(* CODESYS project Portal_robot.project

Project tree, tasks and I/O mapping:
  Device : LicOS-PAC-MC522, Unionscience Technology Group Co.,Ltd, order no. 50080156/50080256, version 3.5.18.50
      unmapped channels: ErrCode
    application Application
      libraries: Standard, 3.5.18.0 (System); CmpBitmapPool, * (System); ModbusFB, 4.3.0.0 (3S - Smart Software Solutions GmbH)
      task MainTask (cyclic, interval t#4ms, priority 0) calls PLC_PRG
      task StatisticTask (freewheeling, priority 3) calls STATISTIC
      task SoftMotion_PlanningTask (cyclic, interval t#2ms, priority 1) calls nothing
      image pool HMI_Image
      axis group AXIS_GROUP_XYZ: TRAFO.Kin_Gantry3, axes X, Y, Z
      Symbols
      FB/
        function block FB_MAGAZINE [ST]: FindBlank, UpdateErrorView, FindFreeSlot, UpdateTypeStatus
        function block FB_TWO_PALLET_SIMULATION [ST]
        function block FB_MOTION_MANAGER [ST]: UpdateErrorView
        function block FB_ALARM_MANAGER [ST]: DeactivateEvent, GetAlarmEffect, AddEvent, UpdateSource
        function block FB_SIMULATION_DYNAMIC_LIMITS [ST]
        function block FB_AXIS [ST]: UpdateErrorView
        function block FB_ALARM_HORN [ST]
        function F_GEOMETRY_EVENT [ST]
        function block FB_GRIPPER_SIMULATION [ST]: UpdateErrorView
        function block FB_MACHINE [ST]: UpdateErrorView
        function block FB_AXIS_GROUP [ST]: UpdateErrorView
        function block FB_GEOMETRY_CONTROL_SIMULATION [ST]
        function block FB_POINT_MANAGER [ST]: UpdateErrorView
        function block FB_ROBOT_MODBUS [ST]
        function block FB_DI_FILTER [ST]
        function block FB_GEOMETRY_CONTROL [ST]
        _ARCHIVE_LEGACY_MULTI_TYPE_HELPERS/
          function block FB_MAGAZINE_RETURN_BLANK_LEGACY [ST]
          function block FB_MAGAZINE_MULTI_TYPE_MAP_LEGACY [ST]
        FB_FAULT_INJECTOR/
          function block FB_ROBOT_FAULT_INJECTOR [ST]
          function block FB_MAGAZINE_FAULT_INJECTOR [ST]
          function block FB_CELL_SAFETY_FAULT_INJECTOR [ST]
          function block FB_CELL_FAULT_INJECTOR [ST]
          function block FB_AXIS_GROUP_FAULT_INJECTOR [ST]
          function block FB_POINT_FAULT_INJECTOR [ST]
          function block FB_GRIPPER_FAULT_INJECTOR [ST]
          function block FB_MACHINE_FAULT_INJECTOR [ST]
          function block FB_AXIS_FAULT_INJECTOR [ST]
        function block FB_ROBOT [ST]: UpdateErrorView
        _ARCHIVE_LEGACY_CELL_MANAGER/
          function block FB_CELL_MANAGER_LEGACY [ST]: UpdateErrorView, SelectMachine
        function F_GEOMETRY_SELECT_STATION [ST]
        function block FB_TWO_PALLET [ST]: IsSignalConfigurationValid, UpdateErrorView
        FB_STATISTIC/
          function block FB_CALCULATE [ST]
          function block FB_STATISTIC [ST]
        function block FB_MACHINE_SIMULATION [ST]: UpdateErrorView
        FB_MULTI_TYPE/
          function block FB_MULTI_TYPE_CONFIG_MANAGER [ST]: ApplyDistribution, RaiseWarning
        function F_GEOMETRY_FIRST_CALL [ST]
        FB_CELL_MANAGER/
          function block FB_CELL_MANAGER [ST]: IsMachineEligible, RaisePayloadRouteWarning, RunGeometryRoute, IsMachineCompatible, SelectMachineBeforeTake, PlanGeometry, UpdateErrorView, SelectMachineForUnload, UpdateGeometryWait, SelectMachineForHeldBlank, CanReturnHeldBlank
        function block FB_CELL_SAFETY [ST]: RaiseWarning
        function F_GEOMETRY_TAKE_DETAIL [ST]
      program PLC_PRG [ST]: ReadHmiInputs, ResetIoEmergencyStop, ReadHmiCommands, RunRobotModbus, RunRobot, RunTwoPallet, RunCellControl, RunTestControl, RunSignalTower, AppendIoEvent, RunMagazine, RunTwoPalletAxis, ReadIoEmergencyStop, RunMotion, RunGeometryControl, RunMachines, ApplyIoOutputOverrides, RunAlarms, ReadPhysicalInputs, RecordIoDiagnostics, PublishGeometryControl, SetApplicationDefaults, RunSafety, ReadIoOverrides, PublishHmi, IsHmiCommandFresh, WritePhysicalOutputs
      ST/
        ST_GRIPPER/
          data type E_GRIPPER_STATE
          data type ST_GRIPPER_DIAG
          data type ST_GRIPPER_COMMAND
          data type ST_GRIPPER_STATUS
          data type ST_GRIPPER_FAULT_REQUEST
          data type ST_GRIPPER_ERRORS
          data type ST_GRIPPER_ERROR
        ST_MULTI_TYPE/
          data type ST_MULTI_TYPE_CONFIG_STATUS
          data type ST_MULTI_TYPE_COMMAND
          data type ST_MULTI_TYPE_CONFIG
          data type ST_MULTI_TYPE_HMI
        ST_ALARM/
          data type ST_ALARM_EVENT
          data type E_ALARM_EFFECT
          data type ST_ALARM_STATUS
          data type ST_ALARM_COMMAND
          data type E_ALARM_SEVERITY
          data type ST_WARNING_EVENT
          data type ST_ALARM_SOURCE_DATA
          data type E_ALARM_SOURCE
        ST_HMI/
          data type ST_PHYSICAL_IO_EVENT
          data type ST_AXIS_HMI_COMMAND
          data type ST_HMI
          data type ST_ROBOT_HMI_STATUS
          data type E_HMI_MANUAL_REJECT
          data type ST_AXIS_HMI_STATUS
        ST_POINT/
          data type ST_POINT
          data type E_POINT_NAME
        ST_ROBOT/
          data type ST_ROBOT_MODBUS_CONFIG
          data type ST_ROBOT_STATUS
          data type E_ROBOT_MODBUS_EXECUTION_STATE
          data type E_ROBOT_MODBUS_CLIENT_STATE
          data type ST_ROBOT_MODBUS_STATUS
          data type ST_ROBOT_FAULT_STATUS
          data type ST_ROBOT_ERRORS
          data type ST_ROBOT_FAULT_REQUEST
          data type ST_ROBOT_DIAG
          data type E_ROBOT_STATE
          data type ST_ROBOT_COMMAND
          data type ST_ROBOT_ERROR
          data type E_ROBOT_ACTION
          data type E_ROBOT_CONTROL_MODE
        ST_CELL/
          data type ST_CELL_DIAG
          data type ST_CELL_ERROR
          data type ST_CELL_SAFETY_DIAG
          data type ST_CELL_SAFETY_ERRORS
          data type ST_CELL_CYCLE_STATUS
          data type ST_ENCLOSURE_DOOR_STATUS
          data type ST_CELL_ERRORS
          data type ST_CELL_COMMAND
          data type ST_BUTTON_STATION_IO_STATUS
          data type E_CELL_MANAGER_STATE
          data type ST_CELL_FAULT_REQUEST
          data type ST_CONTROL_CABINET_IO_STATUS
          data type ST_CELL_STATUS
          data type ST_CELL_SAFETY_STATUS
          data type ST_MPG_IO_STATUS
          data type ST_CELL_SAFETY_FAULT_REQUEST
          data type E_CELL_STATE
        ST_TEST/
          data type ST_TEST_OBSERVABILITY
          data type ST_TEST_SCENARIO_BUFFER
          data type E_CELL_TEST_ENVIRONMENT
          data type E_TEST_SPEED_PROFILE
        ST_AXIS_GROUP/
          data type ST_AXIS_GROUP_ERROR
          data type ST_AXIS_GROUP_ERRORS
          data type ST_AXIS_GROUP_COMMANDS
          data type ST_AXIS_GROUP
          data type ST_AXIS_GROUP_TIMEOUTS
          data type ST_AXIS_GROUP_FAULT_REQUEST
          data type ST_AXIS_GROUP_MOTION_PARAMS
          data type E_AXIS_GROUP_POWER_MODE
          data type E_AXIS_GROUP_STATE
          data type ST_AXIS_GROUP_STATUS
          data type E_MOTION_RESET_STATE
          data type ST_AXIS_GROUP_DIAGNOSTICS
        ST_MOTION_MANAGER/
          data type ST_MOTION_MANAGER_DIAG
          data type ST_MOTION_MANAGER_ERROR
          data type ST_MOTION_MANAGER_COMMAND
          data type E_MOTION_MANAGER_STATE
          data type ST_MOTION_MANAGER
          data type ST_MOTION_MANAGER_ERRORS
          data type ST_MOTION_MANAGER_STATUS
        ST_POINT_MANAGER/
          data type ST_POINT_MANAGER_DIAG
          data type ST_POINT_FAULT_REQUEST
          data type ST_POINT_MANAGER_COMMAND
          data type E_POINT_MANAGER_STATE
          data type ST_POINT_MANAGER_ERRORS
          data type ST_POINT_MANAGER
          data type ST_POINT_MANAGER_ERROR
          data type ST_POINT_MANAGER_STATUS
        ST_MACHINE/
          data type ST_MACHINE_COMMAND
          data type E_PART_TYPE
          data type E_PART_STATE
          data type ST_MACHINE_SIM_ERROR
          data type ST_MACHINE_SIM_ERRORS
          data type ST_MACHINE_ERRORS
          data type ST_MACHINE_POINTS
          data type E_MACHINE_OPERATION
          data type ST_MACHINE_SIM_DIAG
          data type ST_MACHINE_ERROR
          data type ST_MACHINE_RECIPE
          data type ST_MACHINE_TIMEOUTS
          data type E_MACHINE_STATE
          data type ST_MACHINE_DIAG
          data type ST_MACHINE_IO_COMMAND
          data type ST_MACHINE_FAULT_REQUEST
          data type ST_MACHINE_IO_STATUS
          data type E_MACHINE_POINTS
          data type ST_MACHINE_PUBLIC
        ST_STATISTIC/
          data type ST_STATISTIC
          data type ST_STATISTIC_MACHINE
          data type ST_STATISTIC_ROBOT
        ST_GEOMETRY_CONTROL/
          data type ST_GEOMETRY_CALL
          data type ST_GEOMETRY_REQUEST
          data type ST_GEOMETRY_MEMORY
          data type ST_GEOMETRY_STATUS
          data type ST_GEOMETRY_CONFIG
          data type ST_GEOMETRY_SIGNALS
          data type ST_GEOMETRY_EVENT
        ST_MAGAZINE/
          data type ST_TWO_PALLET_ERROR
          data type ST_MAGAZINE_ERROR
          data type ST_MAGAZINE_TYPE_STATUS
          data type ST_MAGAZINE_STATUS
          data type ST_TWO_PALLET_INPUT
          data type ST_TWO_PALLET_ERRORS
          data type ST_MAGAZINE_DIAG
          data type ST_TWO_PALLET_COMMAND
          data type ST_MAGAZINE_FAULT_REQUEST
          data type ST_TWO_PALLET_DIAG
          data type ST_MAGAZINE_ERRORS
          data type ST_MAGAZINE_COMMAND
          data type E_MAGAZINE_STATE
          ST_DETAIL/
            data type E_DETAIL_TYPE
            data type ST_DETAIL
          data type E_TWO_PALLET_STATE
          data type ST_TWO_PALLET_CONFIG
          data type ST_MAGAZINE_HMI_COMMAND
          data type ST_TWO_PALLET_STATUS
          data type ST_TWO_PALLET_STORE
          data type E_MAGAZINE_OPERATION
          data type ST_MAGAZINE_INVENTORY
          data type ST_TWO_PALLET_REQUEST
          data type ST_TWO_PALLET_OUTPUT
        ST_AXIS/
          data type ST_AXIS_DIAGNOSTICS
          data type ST_AXIS_MOTION_PARAMS
          data type E_AXIS_STATE
          data type ST_AXIS_TIMEOUTS
          data type ST_AXIS_ERROR_CODES
          data type ST_AXIS_FAULT_REQUEST
          data type ST_AXIS
          data type ST_AXIS_STATUS
          data type ST_AXIS_ERROR
          data type ST_AXIS_COMMANDS
        ST_FAULT_INJECTOR/
          data type ST_FAULT_INJECTION_STATUS
      program STATISTIC [ST]
      GVL/
        global variables GVL_MAGAZINE
        global variables GVL_ROBOT
        global variables GVL_MAGAZINE_AXIS
        global variables GVL_MACHINE
        global variables GVL_POINT_MANAGER
        global variables GVL_HMI
        global variables GVL_AXIS_GROUP
        global variables GVL_ROBOT_MODBUS
        global variables GVL_CELL_CONTROL
        global variables GVL_CELL_MANAGER
        global variables GVL_POINT
        global variables GVL_ALARM
        global variables GVL_STATISTIC
        global variables GVL_ROBOT_MODBUS_RETAIN
        global variables GVL_CELL_SAFETY_IO
        global variables GVL_GEOMETRY_CONTROL
        global variables GVL_TEST_IO
        global variables GVL_CELL_SETTINGS
        global variables GVL_DETAIL
        global variables GVL_AXIS
        global variables GVL_MULTI_TYPE
        global variables GVL_MOTION_MANAGER
        global variables GVL_PHYSICAL_IO
        global variables GVL_TWO_PALLET
    SoftMotion General Axis Pool
      Z : SM_Drive_Virtual, 3S - Smart Software Solutions GmbH, order no. 1805, version 4.0.0.0
          settings: wDriveID = 0; fSWMaxVelocity = 3300; fSWMaxAcceleration = 12000; fSWMaxDeceleration = 12000; fSWMaxJerk = 100000; fSWLimitPositive = 10000.0; fSWLimitNegative = -1000.0; bSWLimitEnable = TRUE
      X : SM_Drive_Virtual, 3S - Smart Software Solutions GmbH, order no. 1805, version 4.0.0.0
          settings: fSWMaxVelocity = 3300; fSWMaxAcceleration = 12000; fSWMaxDeceleration = 12000; fSWMaxJerk = 100000; fSWLimitPositive = 13000.0; fSWLimitNegative = -1000.0; bSWLimitEnable = TRUE
      Y : SM_Drive_Virtual, 3S - Smart Software Solutions GmbH, order no. 1805, version 4.0.0.0
          settings: wDriveID = 2; fSWMaxVelocity = 3300; fSWMaxAcceleration = 12000; fSWMaxDeceleration = 12000; fSWMaxJerk = 100000; fSWLimitPositive = 10000.0; fSWLimitNegative = -1000.0; bSWLimitEnable = TRUE
      Magazine_1 : SM_Drive_Virtual, 3S - Smart Software Solutions GmbH, order no. 1805, version 4.0.0.0
          settings: wDriveID = 3; fSWMaxVelocity = 3300; fSWMaxAcceleration = 12000; fSWMaxDeceleration = 12000; fSWMaxJerk = 100000; fSWLimitPositive = 13000.0; fSWLimitNegative = -1000.0; bSWLimitEnable = TRUE
      Magazine_2 : SM_Drive_Virtual, 3S - Smart Software Solutions GmbH, order no. 1805, version 4.0.0.0
          settings: wDriveID = 4; fSWMaxVelocity = 3300; fSWMaxAcceleration = 12000; fSWMaxDeceleration = 12000; fSWMaxJerk = 100000; fSWLimitPositive = 13000.0; fSWLimitNegative = -1000.0; bSWLimitEnable = TRUE
    LicOS_MQTT : Mqtt Brok Sub Pub, Unionscience Technology Group Co.,Ltd, order no. 50010000, version 02.00.00.01
    LicOS_MTCP : ModbusTCP Device, Unionscience Technology Group Co.,Ltd, order no. 50011000, version 03.00.00.01
    LicOS_MUDP : ModbusUDP Device, Unionscience Technology Group Co.,Ltd, order no. 50011100, version 03.00.00.01
    LicOS_MRTU : ModbusRTU Device, Unionscience Technology Group Co.,Ltd, order no. 50012000, version 03.00.00.01
    LicOS_NETC : UDP/TCP NetComm, Unionscience Technology Group Co.,Ltd, order no. 50015000, version 01.00.00.01
    LicOS_INTM : Interrupt Cfg Module, Unionscience Technology Group Co.,Ltd, order no. 20110000, version 01.00.00.01
        unmapped channels: ErrCode
  libraries: VisuSymbols, 4.1.0.0 (System)
  text list GlobalTextList
*)

// Device/Application/ST/ST_CELL/ST_CELL_DIAG
TYPE ST_CELL_DIAG :
STRUCT
	eState : E_CELL_STATE; // Текущее состояние автомата ячейки
	stWarning : ST_WARNING_EVENT; // Последнее предупреждение менеджера ячейки
END_STRUCT
END_TYPE

// Device/Application/ST/ST_ROBOT/ST_ROBOT_MODBUS_CONFIG
TYPE ST_ROBOT_MODBUS_CONFIG :
STRUCT
	aIpAddress        : ARRAY [0..3] OF BYTE; // IPv4 контроллера робота
	uiPort            : UINT := UINT#502; // TCP-порт Modbus
	uiUnitId          : UINT := UINT#1; // Unit ID в Modbus TCP
	tResponseTimeout  : TIME := T#500MS; // Ожидание ответа FC03/FC16
	tPollInterval     : TIME := T#50MS; // Период чтения обратной связи
	tHeartbeatTimeout : TIME := T#2S; // Максимальная пауза heartbeat робота
	tCommandTimeout   : TIME := T#600S; // Предельная длительность одной команды
END_STRUCT
END_TYPE

// Device/Application/ST/ST_MOTION_MANAGER/ST_MOTION_MANAGER_DIAG
TYPE ST_MOTION_MANAGER_DIAG :
STRUCT
	eState : E_MOTION_MANAGER_STATE; // Текущее состояние автомата движения
	stWarning : ST_WARNING_EVENT; // Последнее предупреждение менеджера движения
END_STRUCT
END_TYPE

// Device/Application/ST/ST_CELL/ST_CELL_ERROR
TYPE ST_CELL_ERROR :
STRUCT
	BOTH_GRIPPERS_OCCUPIED : BOOL; // Совместимый бит: диагностическая ошибка согласованности захватов
	ROBOT_ERROR            : BOOL; // Ошибка робота во время автоматического цикла
	MAGAZINE_ERROR         : BOOL; // Ошибка магазина во время операции
	MACHINE_ERROR          : BOOL; // Ошибка станка во время обслуживания
	GLOBAL_STOP            : BOOL; // Получена глобальная ошибка ячейки
END_STRUCT
END_TYPE

// Device/Application/ST/ST_POINT_MANAGER/ST_POINT_MANAGER_DIAG
TYPE ST_POINT_MANAGER_DIAG :
STRUCT
	eState       : E_POINT_MANAGER_STATE; // Текущее состояние автомата
	lrX_MinLimit : LREAL; // Минимально допустимая координата X
	lrY_MinLimit : LREAL; // Минимально допустимая координата Y
	lrZ_MinLimit : LREAL; // Минимально допустимая координата Z
	lrX_MaxLimit : LREAL; // Максимально допустимая координата X
	lrY_MaxLimit : LREAL; // Максимально допустимая координата Y
	lrZ_MaxLimit : LREAL; // Максимально допустимая координата Z
	xXLimitValid : BOOL; // Software limits оси X включены и образуют корректный диапазон
	xYLimitValid : BOOL; // Software limits оси Y включены и образуют корректный диапазон
	xZLimitValid : BOOL; // Software limits оси Z включены и образуют корректный диапазон
	stWarning    : ST_WARNING_EVENT; // Последнее предупреждение менеджера точек
END_STRUCT
END_TYPE

// Device/Application/ST/ST_CELL/ST_CELL_SAFETY_DIAG
TYPE ST_CELL_SAFETY_DIAG :
STRUCT
	stWarning : ST_WARNING_EVENT; // Отклонённые попытки открытия и сброса реле
END_STRUCT
END_TYPE

// Device/Application/ST/ST_CELL/ST_CELL_SAFETY_ERRORS
TYPE ST_CELL_SAFETY_ERRORS :
STRUCT
	dwErrorActive : DWORD; // Текущие отдельные Safety-причины
	dwErrorLast   : DWORD; // Последняя ненулевая маска для диагностики
	dwAlarmActive : DWORD; // Собственные аварии источника для общего журнала
END_STRUCT
END_TYPE

// Device/Application/ST/ST_CELL/ST_CELL_CYCLE_STATUS
TYPE ST_CELL_CYCLE_STATUS :
STRUCT
	eState              : E_CELL_MANAGER_STATE; // Состояние универсального автомата ячейки
	uiSelectedMachine   : UINT; // Зафиксированный целевой станок
	uiSelectedType      : UINT; // Тип заготовки текущего маршрута
	uiBlankPayloadType  : UINT; // Тип заготовки в первом захвате
	uiDetailPayloadType : UINT; // Тип готовой детали во втором захвате
	iTakeSlot           : SINT; // Зарезервированный слот взятия
	iPutSlot            : SINT; // Зарезервированный слот укладки
	xReturningBlank     : BOOL; // Выполняется возврат заготовки
	axMachineStartPending: ARRAY [1..3] OF BOOL; // Запуск нового цикла ещё подтверждается станком
	auiBlankCount       : ARRAY [1..3] OF UINT; // Заготовки по типам
	auiDetailCount      : ARRAY [1..3] OF UINT; // Готовые детали по типам
	auiFreeCount        : ARRAY [1..3] OF UINT; // Свободные слоты по типам
END_STRUCT
END_TYPE

// Device/Application/ST/ST_TEST/ST_TEST_OBSERVABILITY
TYPE ST_TEST_OBSERVABILITY :
STRUCT
	udiAppliedScenarioSeq : UDINT;
	uiCellState : UINT;
	uiRobotState : UINT;
	uiRobotAction : UINT;
	uiRobotPoint : UINT;
	uiActiveMagazine : UINT;
	uiMagazineState : UINT;
	uiMagazineOperation : UINT;
	uiTakeSlot : UINT;
	uiPutSlot : UINT;
	auiMachineState : ARRAY [1..3] OF UINT;
	auiMachineOperation : ARRAY [1..3] OF UINT;
	uiSelectedMachine : UINT;
	uiSelectedType : UINT;
	uiErrorSource : UINT;
	dwErrorCode : DWORD;
END_STRUCT
END_TYPE

// Device/Application/ST/ST_MACHINE/ST_MACHINE_COMMAND
TYPE ST_MACHINE_COMMAND :
STRUCT
	stIo    : ST_MACHINE_IO_COMMAND; // Команды исполнительным механизмам станка
	stRobot : ST_ROBOT_COMMAND; // Команда роботу от алгоритма станка
END_STRUCT
END_TYPE

// Device/Application/ST/ST_MACHINE/E_PART_TYPE
{attribute 'qualified_only'}
{attribute 'strict'}
TYPE E_PART_TYPE :
(
	UNKNOWN,
	DETAIL,
	PART
);
END_TYPE

// Device/Application/ST/ST_MACHINE/E_PART_STATE
{attribute 'qualified_only'}
{attribute 'strict'}
TYPE E_PART_STATE :
(
	UNKNOWN := 0,
    EMPTY   := 1,
    LOADED  := 2
);
END_TYPE

// Device/Application/ST/ST_POINT_MANAGER/ST_POINT_FAULT_REQUEST
TYPE ST_POINT_FAULT_REQUEST :
STRUCT
	xEnabled        : BOOL; // Глобальное разрешение диагностической инъекции
	xXOutOfLimit    : BOOL; // Импульс проверки точки с недопустимой координатой X
	xYOutOfLimit    : BOOL; // Импульс проверки точки с недопустимой координатой Y
	xZOutOfLimit    : BOOL; // Импульс проверки точки с недопустимой координатой Z
	xInvalidVelocity: BOOL; // Импульс проверки точки с недопустимой скоростью
END_STRUCT
END_TYPE

// Device/Application/ST/ST_ROBOT/ST_ROBOT_STATUS
TYPE ST_ROBOT_STATUS :
STRUCT
	xBusy             : BOOL; // Робот выполняет команду
	xDone             : BOOL; // Команда завершена
	xError            : BOOL; // Робот находится в ошибке
	xExternalError    : BOOL; // Робот остановлен ошибкой зависимого блока
	xPowerAllowed     : BOOL; // Кнопка включения или отключения приводов доступна
	xStopAllowed      : BOOL; // Кнопка контролируемой остановки доступна
	xResetAllowed     : BOOL; // Кнопка сброса ошибок робота и приводов доступна
	eCurrentPoint     : E_POINT_NAME; // Последняя достигнутая точка
	uiMagazineContext : UINT; // 0 вне рабочей зоны; 1..2 — магазин, в рабочей зоне которого находится робот
	xBlankAvailable   : BOOL; // В первом захвате находится заготовка
	xDetailAvailable  : BOOL; // Во втором захвате находится готовая деталь
	uiBlankPayloadType  : UINT; // Фактический тип заготовки, 0 — неизвестно
	uiDetailPayloadType : UINT; // Фактический тип детали, 0 — неизвестно
	xGripper1Open     : BOOL; // Первый захват открыт
	xGripper1Closed   : BOOL; // Первый захват закрыт
	xGripper2Open     : BOOL; // Второй захват открыт
	xGripper2Closed   : BOOL; // Второй захват закрыт
	xRotatedToBlank   : BOOL; // Захват повёрнут к заготовке
	xRotatedToDetail  : BOOL; // Захват повёрнут к готовой детали
END_STRUCT
END_TYPE

// Device/Application/ST/ST_ROBOT/E_ROBOT_MODBUS_EXECUTION_STATE
{attribute 'qualified_only'}
{attribute 'strict'}
TYPE E_ROBOT_MODBUS_EXECUTION_STATE :
(
	IDLE := 0,
	ACCEPTED := 1,
	BUSY := 2,
	DONE := 3,
	ERROR := 4,
	STOPPED := 5
);
END_TYPE

// Device/Application/ST/ST_CELL/ST_ENCLOSURE_DOOR_STATUS
TYPE ST_ENCLOSURE_DOOR_STATUS :
STRUCT
	xLocked        : BOOL; // Обратная связь замка: TRUE — замок закрыт
	xUnlockAllowed : BOOL; // PLC разрешает открыть замок
	xUnlockOutput  : BOOL; // Фактическая команда открытия замка
END_STRUCT
END_TYPE

// Device/Application/ST/ST_ROBOT/E_ROBOT_MODBUS_CLIENT_STATE
{attribute 'qualified_only'}
{attribute 'strict'}
TYPE E_ROBOT_MODBUS_CLIENT_STATE :
(
	DISABLED,
	CONNECTING,
	INITIAL_READ,
	INITIAL_READ_RELEASE,
	CLEAR_COMMAND,
	CLEAR_COMMAND_RELEASE,
	READY,
	WRITE_COMMAND,
	WRITE_COMMAND_RELEASE,
	READ_STATUS,
	READ_STATUS_RELEASE,
	RECONNECT_WAIT
);
END_TYPE

// Device/Application/ST/ST_MAGAZINE/ST_TWO_PALLET_ERROR
TYPE ST_TWO_PALLET_ERROR :
STRUCT
	DRIVE_ERROR : BOOL;
	SENSOR_CONTRADICTION : BOOL;
	CYLINDER_TIMEOUT : BOOL;
	MOTION_TIMEOUT : BOOL;
	LOGIC_ERROR : BOOL;
	SEQUENCE_INTERRUPTED : BOOL;
END_STRUCT
END_TYPE

// Device/Application/ST/ST_MOTION_MANAGER/ST_MOTION_MANAGER_ERROR
TYPE ST_MOTION_MANAGER_ERROR :
STRUCT
	POINT_INVALID : BOOL; // Целевая точка не прошла проверку
	GROUP_ERROR   : BOOL; // Группа осей завершила движение с ошибкой
	GLOBAL_STOP   : BOOL; // Получена глобальная ошибка ячейки
	START_TIMEOUT : BOOL; // Истекло ожидание проверки точки или старта группы
END_STRUCT
END_TYPE

// Device/Application/ST/ST_AXIS/ST_AXIS_DIAGNOSTICS
TYPE ST_AXIS_DIAGNOSTICS :
STRUCT
    iStep            : E_AXIS_STATE; // Текущий шаг автомата оси
    iLastErrorStep   : INT; // Шаг, на котором возникла последняя ошибка
    sStepName        : STRING[80]; // Текстовое имя текущего шага
    sWaitReason      : STRING[120]; // Причина ожидания на текущем шаге
    sErrorText       : STRING[120]; // Текст активной ошибки
    sWarningText     : STRING[120]; // Текст активного предупреждения
    stWarning        : ST_WARNING_EVENT; // Последнее предупреждение оси для общего журнала
    tStepElapsed     : TIME; // Время нахождения на текущем шаге
    tStepPreset      : TIME; // Допустимое время текущего шага
    xStepTimeout     : BOOL; // Превышено допустимое время шага
    udiActualErrorID : UDINT; // Код активной ошибки
    udiLastErrorID   : UDINT; // Код последней ошибки
END_STRUCT
END_TYPE

// Device/Application/ST/ST_CELL/ST_CELL_ERRORS
TYPE ST_CELL_ERRORS :
STRUCT
	dwErrorActive : DWORD; // Битовая маска активных ошибок
	dwErrorLast   : DWORD; // Битовая маска последних ошибок
	dwAlarmActive : DWORD; // Собственные аварии менеджера ячейки для общего журнала
	stErrorActive : ST_CELL_ERROR; // Расшифровка активных ошибок
	stErrorLast   : ST_CELL_ERROR; // Расшифровка последних ошибок
END_STRUCT
END_TYPE

// Device/Application/ST/ST_AXIS/ST_AXIS_MOTION_PARAMS
TYPE ST_AXIS_MOTION_PARAMS :
STRUCT
    lrTargetPosition : LREAL; // Целевая абсолютная позиция
    lrDistance       : LREAL; // Дистанция относительного перемещения
    lrHomePosition   : LREAL; // Координата домашней позиции
    lrVelocity       : LREAL; // Скорость движения
    lrAcceleration   : LREAL; // Ускорение
    lrDeceleration   : LREAL; // Замедление
    lrJerk           : LREAL; // Рывок
END_STRUCT
END_TYPE

// Device/Application/ST/ST_ROBOT/ST_ROBOT_MODBUS_STATUS
TYPE ST_ROBOT_MODBUS_STATUS :
STRUCT
	xConfigValid       : BOOL; // Параметры соединения прошли проверку PLC
	xConnected         : BOOL; // TCP-соединение установлено
	xCommunicationAlive: BOOL; // Получена свежая обратная связь и меняется heartbeat
	xStatusFresh       : BOOL; // После подключения успешно прочитан блок 1101..1117
	xControllerOn      : BOOL;
	xAutomaticMode     : BOOL;
	xRemoteEnabled     : BOOL;
	xDrivesEnabled     : BOOL;
	xHomed             : BOOL;
	xEmergencyStop     : BOOL;
	xRobotAlarm        : BOOL;
	xPositionValid     : BOOL;
	xSimulatorActive   : BOOL; // Бит 1108.9: подключён Python-симулятор, а не реальный SC-500
	xReady             : BOOL; // Итоговая готовность, пересчитанная PLC
	xBusy              : BOOL;
	xDone              : BOOL;
	xError             : BOOL; // Ошибка исполнения, робота или транспорта
	xCommandTimeout    : BOOL; // Робот не завершил принятую команду за лимит
	xResetBusy         : BOOL; // Передача Reset и подтверждение его снятия ещё выполняются
	xResetDone         : BOOL; // Reset подтверждён обратной связью и очищенной FC16
	xResetFailed       : BOOL; // Попытка сорвана/истекла; повтор только новым запросом
	uiAckSeq           : UINT;
	uiExecutionState   : UINT;
	uiResultCode       : UINT;
	uiActiveCommand    : UINT;
	uiCurrentPoint     : UINT;
	uiGripperStatus    : UINT;
	uiRobotHeartbeat   : UINT;
	uiStatusWord       : UINT;
	uiAlarmCode        : UINT;
	uiOperationPhase   : UINT;
	uiProtocolVersion  : UINT;
	lrActualX          : LREAL;
	lrActualY          : LREAL;
	lrActualZ          : LREAL;
	udiClientError     : UDINT;
	udiReadError       : UDINT;
	udiWriteError      : UDINT;
END_STRUCT
END_TYPE

// Device/Application/ST/ST_AXIS/E_AXIS_STATE
{attribute 'qualified_only'}
{attribute 'strict'}
TYPE E_AXIS_STATE :
(
	DISABLED,
	POWERING,
	POWERING_DOWN,
	READY,
	JOGGING,
	JOG_DECELERATING,
	HOMING,
	MOVE_ABSOLUTE,
	MOVE_RELATIVE,
	STOPPING,
	STOP_RELEASE,
	ERROR_RESET_MANAGER,
	RESET_AXIS_ERROR,
	RESET_RELEASE,
	RESET_FINISH
);
END_TYPE

// Device/Application/ST/ST_AXIS/ST_AXIS_TIMEOUTS
TYPE ST_AXIS_TIMEOUTS :
STRUCT
	xDisableOnError : BOOL := TRUE; // Отключать привод при логической ошибке
    tPowerFeedbackLossTimeout : TIME := T#500MS; // Потеря силовой готовности при сохраняющемся запросе питания
    tPowerTimeout   : TIME := T#5S; // Время ожидания включения или отключения питания
    tResetTimeout   : TIME := T#5S; // Время ожидания сброса ошибки
    tStopTimeout    : TIME := T#5S; // Время ожидания остановки
    tHomeTimeout    : TIME := T#30S; // Время ожидания поиска домашней позиции
    tMoveTimeout    : TIME := T#15S; // Время ожидания завершения перемещения
END_STRUCT
END_TYPE

// Device/Application/ST/ST_ALARM/ST_ALARM_EVENT
TYPE ST_ALARM_EVENT :
STRUCT
	udiSequence : UDINT; // Уникальный порядковый номер события
	eSeverity   : E_ALARM_SEVERITY; // Уровень события
	eEffect     : E_ALARM_EFFECT; // Фактическое воздействие события в момент фиксации
	eSource     : E_ALARM_SOURCE; // Механизм-источник события
	uiCode      : UINT; // Номер бита ошибки или код предупреждения
	xActive     : BOOL; // Событие ещё активно и требует внимания
END_STRUCT
END_TYPE

// Device/Application/ST/ST_POINT_MANAGER/ST_POINT_MANAGER_COMMAND
TYPE ST_POINT_MANAGER_COMMAND :
STRUCT
	xExecute : BOOL; // Команда проверки заданной точки
END_STRUCT
END_TYPE

// Device/Application/ST/ST_MOTION_MANAGER/ST_MOTION_MANAGER_COMMAND
TYPE ST_MOTION_MANAGER_COMMAND :
STRUCT 
	eTargetPoint : E_POINT_NAME; // Имя целевой точки
	xGlobalError : BOOL; // Глобальная ошибка ячейки
	xExecute     : BOOL; // Команда запуска движения
	xStop        : BOOL; // Штатная операторская остановка без формирования аварии
	xReset       : BOOL; // Команда сброса ошибки
	xMode        : BOOL; // TRUE: Modbus, FALSE: SoftMotion
END_STRUCT
END_TYPE

// Device/Application/ST/ST_AXIS_GROUP/ST_AXIS_GROUP_ERROR
TYPE ST_AXIS_GROUP_ERROR :
STRUCT
	ENABLE_ERROR          : BOOL; // Ошибка MC_GroupEnable
	POWER_ERROR           : BOOL; // Зарезервировано; питание осей контролируют FB_AXIS
	DISABLE_ERROR         : BOOL; // Ошибка MC_GroupDisable
	RESET_ERROR           : BOOL; // Ошибка MC_GroupReset
	MOVE_DIRECT_ERROR     : BOOL; // Ошибка MC_MoveDirectAbsolute
	MOVE_LINEAR_ERROR     : BOOL; // Ошибка MC_MoveLinearAbsolute
	HALT_ERROR            : BOOL; // Ошибка MC_GroupHalt
	STOP_ERROR            : BOOL; // Ошибка MC_GroupStop
	READ_POSITION_ERROR   : BOOL; // Ошибка чтения позиции группы
	READ_STATUS_ERROR     : BOOL; // Ошибка чтения статуса группы
	READ_GROUP_ERROR      : BOOL; // Ошибка чтения кода ошибки группы
	GROUP_ERROR_STOP      : BOOL; // Группа SoftMotion находится в ErrorStop
	SIMULATED_ERROR       : BOOL; // Тестовая ошибка Motion-FB, сформированная эмулятором
	OVERRIDE_ERROR        : BOOL; // Ошибка MC_GroupSetOverride
	STEP_TIMEOUT          : BOOL; // Превышено время выполнения шага
	INVALID_STATE         : BOOL; // Неизвестное состояние автомата
	POWER_PERMIT_READY    : BOOL; // Нет разрешения питания в готовности
	POWER_PERMIT_LOST     : BOOL; // Потеря разрешения питания в движении
END_STRUCT
END_TYPE

// Device/Application/ST/ST_AXIS_GROUP/ST_AXIS_GROUP_ERRORS
TYPE ST_AXIS_GROUP_ERRORS :
STRUCT
	dwMotionErrorLatched  : DWORD; // Защёлкнутые ошибки SoftMotion
	dwLogicalErrorLatched : DWORD; // Защёлкнутые логические ошибки
	dwLogicalErrorNew     : DWORD; // Новые логические ошибки текущего цикла
	dwMotionErrorNew      : DWORD; // Новые ошибки SoftMotion текущего цикла
	dwMotionErrorActive   : DWORD; // Активные ошибки блоков SoftMotion
	dwMotionErrorPrevious : DWORD; // Ошибки SoftMotion предыдущего цикла
	dwMotionErrorLast     : DWORD; // Последняя ненулевая маска SoftMotion
	dwLogicalErrorLast    : DWORD; // Последняя ненулеевая логическая маска
	dwAlarmActive         : DWORD; // Собственные аварии группы для общего журнала
	stErrorActive         : ST_AXIS_GROUP_ERROR; // Расшифровка активных ошибок
	stErrorLast           : ST_AXIS_GROUP_ERROR; // Расшифровка последних ошибок
END_STRUCT
END_TYPE

// Device/Application/ST/ST_CELL/ST_CELL_COMMAND
TYPE ST_CELL_COMMAND :
STRUCT
	stRobot          : ST_ROBOT_COMMAND; // Команда роботу от менеджера ячейки
	uiBlankPayloadType  : UINT; // Тип заготовки в первом захвате
	uiDetailPayloadType : UINT; // Тип готовой детали во втором захвате
	stMagazine       : ST_MAGAZINE_COMMAND; // Команда магазину
	axMachineExecute : ARRAY [1..3] OF BOOL; // Запуск обслуживания выбранного станка
END_STRUCT
END_TYPE

// Device/Application/ST/ST_AXIS/ST_AXIS_ERROR_CODES
TYPE ST_AXIS_ERROR_CODES :
STRUCT
    dwAxisErrorActual     : DWORD; // Текущие ошибки блоков SoftMotion
    dwAxisErrorLatched    : DWORD; // Защёлкнутые ошибки SoftMotion
    dwAxisError           : DWORD; // Общая активная маска ошибок оси
    dwAxisErrorLast       : DWORD; // Последняя ненулевая маска ошибок оси
    dwDriveAxisErrorID    : DWORD; // Код ошибки привода
    dwLogicalErrorLatched : DWORD; // Защёлкнутые логические ошибки
    dwLogicalError        : DWORD; // Общая активная маска логических ошибок
    dwLogicalErrorLast    : DWORD; // Последняя ненулевая маска логических ошибок
    dwWarningLatched      : DWORD; // Защёлкнутые предупреждения
    dwWarning             : DWORD; // Активные предупреждения
    dwAllError            : DWORD; // Сводная маска ошибок
    dwAlarmActive         : DWORD; // Собственные аварии оси для общего журнала
    stErrorActive         : ST_AXIS_ERROR; // Расшифровка активных ошибок
    stErrorLast           : ST_AXIS_ERROR; // Расшифровка последних ошибок
END_STRUCT
END_TYPE

// Device/Application/ST/ST_MAGAZINE/ST_MAGAZINE_ERROR
TYPE ST_MAGAZINE_ERROR :
STRUCT
	WRONG_OPERATION : BOOL; // Операция не может быть выбрана
	NO_BLANK        : BOOL; // В магазине нет доступной заготовки
	NO_FREE_SLOT    : BOOL; // В магазине нет свободного слота
	INVALID_SLOT    : BOOL; // Номер слота находится вне матрицы
	SLOT_CONTENT    : BOOL; // Содержимое выбранного слота не соответствует операции
	ROBOT_ERROR     : BOOL; // Робот завершил команду с ошибкой
	GLOBAL_STOP     : BOOL; // Получена глобальная ошибка ячейки
	GEOMETRY_ERROR  : BOOL; // Геометрия магазина задана неверно
END_STRUCT
END_TYPE

// Device/Application/ST/ST_GRIPPER/E_GRIPPER_STATE
{attribute 'qualified_only'}
{attribute 'strict'}
TYPE E_GRIPPER_STATE :
(
	IDLE,
    EXECUTE,
    DONE,
    ERROR
);
END_TYPE

// Device/Application/ST/ST_ALARM/E_ALARM_EFFECT
TYPE E_ALARM_EFFECT :
(
	GLOBAL_STOP, // Аварийный останов всей ячейки
	ROBOT_STOP, // Останов робота и текущего взаимодействия с оборудованием
	EQUIPMENT_STOP, // Останов только владельца аварии
	WARNING // Информационное предупреждение без останова
);
END_TYPE

// Device/Application/ST/ST_ROBOT/ST_ROBOT_FAULT_STATUS
TYPE ST_ROBOT_FAULT_STATUS :
STRUCT
	stRobot   : ST_FAULT_INJECTION_STATUS; // Локальная ошибка автомата робота
	stGripper : ST_FAULT_INJECTION_STATUS; // Неисправности виртуального захвата
	stPoint   : ST_FAULT_INJECTION_STATUS; // Ошибки проверки точки движения
END_STRUCT
END_TYPE

// Device/Application/ST/ST_ALARM/ST_ALARM_STATUS
TYPE ST_ALARM_STATUS :
STRUCT
	uiActiveAlarmCount   : UINT; // Число активных аварий
	uiActiveWarningCount : UINT; // Число активных предупреждений
	uiActiveEventCount   : UINT; // Общее число активных событий
	uiHistoryCount       : UINT; // Число записей в журнале
	xAlarmActive         : BOOL; // Есть хотя бы одна активная авария
	xWarningActive       : BOOL; // Есть хотя бы одно активное предупреждение
END_STRUCT
END_TYPE

// Device/Application/ST/ST_MAGAZINE/ST_MAGAZINE_TYPE_STATUS
TYPE ST_MAGAZINE_TYPE_STATUS :
STRUCT
	aiBlankSlot    : ARRAY [1..3] OF SINT; // Первая заготовка каждого типа
	aiFreeSlot     : ARRAY [1..3] OF SINT; // Первый свободный слот каждого типа
	auiBlankCount  : ARRAY [1..3] OF UINT; // Количество заготовок каждого типа
	auiDetailCount : ARRAY [1..3] OF UINT; // Количество готовых деталей каждого типа
	auiFreeCount   : ARRAY [1..3] OF UINT; // Количество свободных слотов каждого типа
END_STRUCT
END_TYPE

// Device/Application/ST/ST_CELL/ST_BUTTON_STATION_IO_STATUS
TYPE ST_BUTTON_STATION_IO_STATUS :
STRUCT
	xEmergencyStopPressed : BOOL; // Нормализованный вход: TRUE — грибок нажат
	xButtonPressed        : BOOL; // Нормализованный вход кнопки открытия замка
	xButtonLightOn        : BOOL; // Фактический выход подсветки кнопки
END_STRUCT
END_TYPE

// Device/Application/ST/ST_MACHINE/ST_MACHINE_SIM_ERROR
TYPE ST_MACHINE_SIM_ERROR :
STRUCT
	MACHINE_ALARM : BOOL; // Активна имитация аварии станка
	DOOR_FAULT    : BOOL; // Ошибка механизма двери
	CHUCK_FAULT   : BOOL; // Ошибка механизма патрона
END_STRUCT
END_TYPE

// Device/Application/ST/ST_GRIPPER/ST_GRIPPER_DIAG
TYPE ST_GRIPPER_DIAG :
STRUCT
	eState        : E_GRIPPER_STATE; // Текущее состояние автомата
	eActiveAction : E_ROBOT_ACTION; // Выполняемое действие захвата
	stWarning     : ST_WARNING_EVENT; // Последнее предупреждение захвата
END_STRUCT
END_TYPE

// Device/Application/ST/ST_HMI/ST_PHYSICAL_IO_EVENT
TYPE ST_PHYSICAL_IO_EVENT :
STRUCT
    udiSequence : UDINT;
    uliTimeMs : ULINT; // Монотонное время от старта приложения, без переполнения TIME
    usiDirection : USINT; // 1 DI; 2 DO
    uiIndex : UINT; // DI 1..84; DO 1..50, index из карты I/O
    usiKind : USINT; // 1 клемма DI; 2 вход программы; 3 DO; 4 подмена DI; 5/6 снять DI; 7 ручной DO; 8/9 возврат DO оператором/программе
    xOld : BOOL;
    xNew : BOOL;
END_STRUCT
END_TYPE

// Device/Application/ST/ST_MAGAZINE/ST_MAGAZINE_STATUS
TYPE ST_MAGAZINE_STATUS :
STRUCT
	xEnabled         : BOOL; // Магазин включен в работу
	xDisablePending  : BOOL; // Отключение выполнится после выхода робота и завершения операции
	xPowerAllowed    : BOOL; // Команда включения/отключения может быть принята
	xEnableSequenceAllowed : BOOL; // PLC разрешает ввести подготовленный магазин в автомат
	xEnableCheckRobotReady : BOOL; // Диагностика готовности роботной операции; не блокирует включение
	xEnableCheckRobotReleased : BOOL; // Диагностика положения робота; не блокирует включение
	xEnableCheckNoError : BOOL; // Нет ошибок магазина и глобальных ошибок ячейки
	xEnableCheckContent : BOOL; // Содержимое кассеты допускает полезную операцию
	xEnableCheckGeometry : BOOL; // Матрица содержит от 1 до 120 активных слотов
	xFillAllowed     : BOOL; // Кнопка заполнения магазина заготовками доступна
	xClearAllowed    : BOOL; // Кнопка очистки магазина доступна
	xEditAllowed     : BOOL; // Содержимое разрешено менять только у выключенного магазина
	xPitchEditAllowed : BOOL; // Общий шаг X/Y можно менять только при выключенных обоих магазинах
	xReady 			 : BOOL; // Магазин готов принять команду
	xBusy  			 : BOOL; // Выполняется операция магазина
	xDone  			 : BOOL; // Операция магазина завершена
	xError          : BOOL; // Магазин находится в ошибке
	xRobotStopRequired : BOOL; // Ошибка магазина требует зависимой аварии робота
	xOutBlank        : BOOL; // В магазине не осталось свободных заготовок
	xOutFreeSlot     : BOOL; // В магазине не осталось свободных слотов
	xCanTake         : BOOL; // Операция TAKE доступна по содержимому магазина
	xCanPut          : BOOL; // Операция PUT доступна по содержимому магазина
	xCanChange       : BOOL; // Операция CHANGE доступна по содержимому магазина
	xCanEnable       : BOOL; // Содержимое позволяет взять/положить груз; не блокирует включение
	xFinished        : BOOL; // Палета завершена; защёлка до смены/правки её рабочего содержимого
	udiProducedPartsTotal : UDINT; // Подтверждённые укладки готовой детали с момента запуска PLC
	uiMagazineId    : UINT; // 1 или 2
	iCurrentBlank    : SINT; // Минимальный номер заготовки в матрице
	iCurrentFreeSlot : SINT; // Минимальный номер свободного слота в матрице
	iSelectedBlank   : SINT; // Номер заготовки, выбранной для текущей операции
	iSelectedFreeSlot: SINT; // Номер свободного слота, выбранного для текущей операции
	eGrantedOperation: E_MAGAZINE_OPERATION; // Доступная операция по текущему состоянию магазина
	eActualOperation : E_MAGAZINE_OPERATION; // Выполняемая операция магазина
	stTypeStatus     : ST_MAGAZINE_TYPE_STATUS; // Содержимое кассеты по типам
END_STRUCT
END_TYPE

// Device/Application/ST/ST_MULTI_TYPE/ST_MULTI_TYPE_CONFIG_STATUS
TYPE ST_MULTI_TYPE_CONFIG_STATUS :
STRUCT
	xMagazineConfigAllowed   : BOOL; // Типы и распределение слотов можно менять
	xTypeCountAllowed        : BOOL; // Количество типов можно менять с применением шаблона
	axMachineTypeAllowed     : ARRAY [1..3] OF BOOL; // Назначение типа конкретному станку разрешено
	xConfigurationValid      : BOOL; // Конфигурация пригодна для автоматического цикла
	uiActiveSlotCount        : UINT; // Число слотов активной матрицы
	stWarning                : ST_WARNING_EVENT; // Последняя отклонённая команда конфигурации
END_STRUCT
END_TYPE

// Device/Application/ST/ST_MACHINE/ST_MACHINE_SIM_ERRORS
TYPE ST_MACHINE_SIM_ERRORS :
STRUCT
	dwErrorActive : DWORD; // Битовая маска активных ошибок
	dwErrorLast   : DWORD; // Битовая маска последних ошибок
	stErrorActive : ST_MACHINE_SIM_ERROR; // Расшифровка активных ошибок
	stErrorLast   : ST_MACHINE_SIM_ERROR; // Расшифровка последних ошибок
END_STRUCT
END_TYPE

// Device/Application/ST/ST_MAGAZINE/ST_TWO_PALLET_INPUT
TYPE ST_TWO_PALLET_INPUT :
STRUCT
	xIoMapped : BOOL; // Подтверждается наладчиком после привязки и проверки физических I/O
	xLiftDown : BOOL;
	xLiftUp : BOOL;
	xLockIn : BOOL;
	xLockOut : BOOL;
	xStopIn : BOOL;
	xStopOut : BOOL;
	xLimitNegative : BOOL;
	xLimitPositive : BOOL;
	xHomeSensor : BOOL; // Только датчик каретки, не палет
	xAxisBound : BOOL;
	xPowered : BOOL;
	xHomed : BOOL;
	xStandstill : BOOL;
	xDriveError : BOOL;
	xMotionDone : BOOL;
	lrPosition : LREAL;
END_STRUCT
END_TYPE

// Device/Application/ST/ST_ROBOT/ST_ROBOT_ERRORS
TYPE ST_ROBOT_ERRORS :
STRUCT
	dwErrorActive : DWORD; // Битовая маска активных ошибок
	dwErrorLast   : DWORD; // Битовая маска последних ошибок
	dwAlarmActive : DWORD; // Собственные аварии робота для общего журнала
	stErrorActive : ST_ROBOT_ERROR; // Расшифровка активных ошибок
	stErrorLast   : ST_ROBOT_ERROR; // Расшифровка последних ошибок
END_STRUCT
END_TYPE

// Device/Application/ST/ST_HMI/ST_AXIS_HMI_COMMAND
TYPE ST_AXIS_HMI_COMMAND :
STRUCT
	xJogPositive      : BOOL; // Удерживаемый Jog в положительном направлении
	xJogNegative      : BOOL; // Удерживаемый Jog в отрицательном направлении
	{attribute 'symbol' := 'read'}
	xHome             : BOOL; // Импульс поиска домашней позиции выбранной оси
	{attribute 'symbol' := 'read'}
	xMoveAbsolute     : BOOL; // Импульс абсолютного перемещения к lrTargetPosition
	{attribute 'symbol' := 'read'}
	xMoveRelative     : BOOL; // Импульс относительного перемещения на lrRelativeDistance
	lrTargetPosition  : LREAL; // Целевая абсолютная координата оси
	lrRelativeDistance : LREAL; // Подготовленная дистанция относительного движения
END_STRUCT
END_TYPE

// Device/Application/ST/ST_HMI/ST_HMI
TYPE ST_HMI :
STRUCT
	ActualX : LREAL; // Текущая координата X для существующей визуализации
	ActualY : LREAL; // Текущая координата Y для существующей визуализации
	ActualZ : LREAL; // Текущая координата Z для существующей визуализации
END_STRUCT
END_TYPE

// Device/Application/ST/ST_GEOMETRY_CONTROL/ST_GEOMETRY_CALL
TYPE ST_GEOMETRY_CALL :
STRUCT
	udiId : UDINT; // Не меняется от вызова до результата контроля
	uiMachine : UINT;
	uiProductType : UINT;
	uiStation : UINT; // 0 до автоматического выбора свободного ГК
	xForced : BOOL;
	uiState : UINT; // 1 вызван, 2 в захвате/ожидание, 3 доставка, 4 на ГК, 5 в магазине, 6 отменён, 7 прерван, 8 изъят
	uiReason : UINT; // 1 заняты оба ГК, 2 нет доступного ГК, 3 отключён, 4 авария, 5 перезапуск/неопределённость
	uiMagazine : UINT;
	uiPallet : UINT;
	uiSlot : UINT;
END_STRUCT
END_TYPE

// Device/Application/ST/ST_STATISTIC/ST_STATISTIC
TYPE ST_STATISTIC :
STRUCT
	stMachineStat 		: ST_STATISTIC_MACHINE;
	stRobotStat 		: ST_STATISTIC_ROBOT;
END_STRUCT
END_TYPE

// Device/Application/ST/ST_ROBOT/ST_ROBOT_FAULT_REQUEST
TYPE ST_ROBOT_FAULT_REQUEST :
STRUCT
	xEnabled     : BOOL; // Глобальное разрешение диагностической инъекции
	xWrongAction : BOOL; // Импульс недопустимого действия робота
	stGripper : ST_GRIPPER_FAULT_REQUEST; // Неисправности виртуального захвата
	stPoint   : ST_POINT_FAULT_REQUEST; // Ошибки проверки точки движения
END_STRUCT
END_TYPE

// Device/Application/ST/ST_MACHINE/ST_MACHINE_ERRORS
TYPE ST_MACHINE_ERRORS :
STRUCT
	dwErrorActive : DWORD; // Битовая маска активных ошибок
	dwErrorLast   : DWORD; // Битовая маска последних ошибок
	dwAlarmActive : DWORD; // Собственные аварии станка для общего журнала
	stErrorActive : ST_MACHINE_ERROR; // Расшифровка активных ошибок
	stErrorLast   : ST_MACHINE_ERROR; // Расшифровка последних ошибок
END_STRUCT
END_TYPE

// Device/Application/ST/ST_MAGAZINE/ST_TWO_PALLET_ERRORS
TYPE ST_TWO_PALLET_ERRORS :
STRUCT
	dwErrorActive : DWORD;
	dwErrorLast : DWORD;
	dwAlarmActive : DWORD;
	stErrorActive : ST_TWO_PALLET_ERROR;
	stErrorLast : ST_TWO_PALLET_ERROR;
END_STRUCT
END_TYPE

// Device/Application/ST/ST_ROBOT/ST_ROBOT_DIAG
TYPE ST_ROBOT_DIAG :
STRUCT
	eState        : E_ROBOT_STATE; // Текущее состояние автомата робота
	eActiveAction : E_ROBOT_ACTION; // Выполняемое действие робота
	eActivePoint  : E_POINT_NAME; // Целевая точка текущего движения
	stWarning     : ST_WARNING_EVENT; // Последнее предупреждение робота
END_STRUCT
END_TYPE

// Device/Application/ST/ST_ALARM/ST_ALARM_COMMAND
TYPE ST_ALARM_COMMAND :
STRUCT
	xResetWarnings : BOOL; // Импульс сброса накопленных предупреждений
END_STRUCT
END_TYPE

// Device/Application/ST/ST_MOTION_MANAGER/E_MOTION_MANAGER_STATE
{attribute 'qualified_only'}
{attribute 'strict'}
TYPE E_MOTION_MANAGER_STATE :
(
	IDLE,
	VALIDATE,
	MOTION_SIM,
	MOTION_MODBUS,
	DONE,
	ERROR
);
END_TYPE

// Device/Application/ST/ST_MOTION_MANAGER/ST_MOTION_MANAGER
TYPE ST_MOTION_MANAGER :
STRUCT
	Command : ST_MOTION_MANAGER_COMMAND; // Команды менеджеру движения
	Status  : ST_MOTION_MANAGER_STATUS; // Рабочие статусы менеджера движения
	Diag    : ST_MOTION_MANAGER_DIAG; // Состояние автомата менеджера движения
	Error   : ST_MOTION_MANAGER_ERRORS; // Активные и последние ошибки
END_STRUCT
END_TYPE

// Device/Application/ST/ST_CELL/E_CELL_MANAGER_STATE
{attribute 'qualified_only'}
{attribute 'strict'}
TYPE E_CELL_MANAGER_STATE :
(
	IDLE,
	PLAN_TARGET,
	MAGAZINE_EXECUTE,
	RELEASE_MAGAZINE,
	ROUTE_TO_TARGET,
	RELEASE_ROBOT_COMMAND,
	WAIT_TARGET,
	SERVICE_TARGET,
	SELECT_FALLBACK,
	WAIT_MAGAZINE,
	ERROR,
	MACHINE_FAULT_STOP,
	PRESTART_IDENTIFY,
	WAIT_GRIPPER1_CONTENT,
	WAIT_GRIPPER1_TYPE,
	WAIT_GRIPPER2_CONTENT,
	WAIT_GRIPPER2_TYPE,
	WAIT_START_MACHINE,
	TEST_ABORT_STOP,
	GEOMETRY_WAIT_FREE,
	GEOMETRY_DELIVER,
	GEOMETRY_RELEASE_COMMAND
);
END_TYPE

// Device/Application/ST/ST_HMI/ST_ROBOT_HMI_STATUS
TYPE ST_ROBOT_HMI_STATUS :
STRUCT
	xDrivesPowered       : BOOL; // Все три привода фактически включены
	xDrivesOff           : BOOL; // Все три привода и группа фактически отключены
	xPowerTransitionActive : BOOL; // Выполняется последовательность включения или отключения
	xDrivesEnableAllowed : BOOL; // PLC разрешает включение приводов
	xDrivesDisableAllowed : BOOL; // PLC разрешает отключение приводов
	xResetAllowed        : BOOL; // PLC разрешает команду сброса ручного управления
	xStopAllowed         : BOOL; // PLC разрешает контролируемую остановку
	xPointsAllowed        : BOOL; // PLC разрешает переход к именованной точке
	xGripperAllowed       : BOOL; // PLC разрешает действие захвата
	xGripper1OpenAllowed  : BOOL;
	xGripper1CloseAllowed : BOOL;
	xGripper2OpenAllowed  : BOOL;
	xGripper2CloseAllowed : BOOL;
	xRotateToBlankAllowed : BOOL;
	xRotateToDetailAllowed : BOOL;
	xCommandBusy          : BOOL;
	uiActiveAction        : UINT;
	uiActivePoint         : UINT;
	eRejectReason         : E_HMI_MANUAL_REJECT; // Числовая причина недоступности команды
END_STRUCT
END_TYPE

// Device/Application/ST/ST_GRIPPER/ST_GRIPPER_COMMAND
TYPE ST_GRIPPER_COMMAND :
STRUCT
	xExecute : BOOL; // Команда запуска действия
	xReset   : BOOL; // Команда сброса ошибки
	eAction  : E_ROBOT_ACTION; // Требуемое действие захвата
	// Дискретный контракт исполнительных механизмов. Каждый BOOL задаёт
	// состояние своего механизма: 0 — закрыть/к заготовке, 1 — открыть/к детали.
	xGripper1Open   : BOOL; // Захват 1: 0 закрыть, 1 открыть
	xGripper2Open   : BOOL; // Захват 2: 0 закрыть, 1 открыть
	xRotateToDetail : BOOL; // Поворот: 0 к заготовке, 1 к детали
END_STRUCT
END_TYPE

// Device/Application/ST/ST_GRIPPER/ST_GRIPPER_STATUS
TYPE ST_GRIPPER_STATUS  :
STRUCT
	xBusy            : BOOL; // Выполняется действие захвата
	xDone            : BOOL; // Действие завершено
	xError           : BOOL; // Захват находится в ошибке
	xGripper1Open    : BOOL; // Первый захват открыт
	xGripper1Closed  : BOOL; // Первый захват закрыт
	xGripper2Open    : BOOL; // Второй захват открыт
	xGripper2Closed  : BOOL; // Второй захват закрыт
	xRotatedToBlank  : BOOL; // Захват повёрнут к заготовке
	xRotatedToDetail : BOOL; // Захват повёрнут к детали
END_STRUCT
END_TYPE

// Device/Application/ST/ST_CELL/ST_CELL_FAULT_REQUEST
TYPE ST_CELL_FAULT_REQUEST :
STRUCT
	xEnabled      : BOOL; // Глобальное разрешение диагностической инъекции
	xBothGrippers : BOOL; // Совместимый диагностический импульс ошибки согласованности захватов
END_STRUCT
END_TYPE

// Device/Application/ST/ST_MACHINE/ST_MACHINE_POINTS
TYPE ST_MACHINE_POINTS :
STRUCT
	eNone          : E_POINT_NAME; // Пустое имя точки
	eAbove         : E_POINT_NAME; // Точка над рабочей зоной станка
	eInside        : E_POINT_NAME; // Точка внутри рабочей зоны станка
	eChuckApproach : E_POINT_NAME; // Точка подхода к патрону
	eChuck         : E_POINT_NAME; // Рабочая точка патрона
END_STRUCT
END_TYPE

// Device/Application/ST/ST_GEOMETRY_CONTROL/ST_GEOMETRY_REQUEST
TYPE ST_GEOMETRY_REQUEST :
STRUCT
	uiAction : UINT; // 1 Enable, 2 Disable, 3 Confirm, 4 Reject, 5 ManualRun, 6 Stop, 7 RemoveSimulation, 8 Call, 9 Auto, 10 Period, 11 Config, 12 Cancel, 13 Capture, 14 SimAlarm, 15 SimAlarmClear, 16 CellSettings
	uiStation : UINT;
	uiMachine : UINT;
	udiValue : UDINT;
	Config : ST_GEOMETRY_CONFIG;
END_STRUCT
END_TYPE

// Device/Application/ST/ST_MAGAZINE/ST_MAGAZINE_DIAG
TYPE ST_MAGAZINE_DIAG :
STRUCT
	eState : E_MAGAZINE_STATE := E_MAGAZINE_STATE.DISABLED; // Текущее состояние автомата магазина
	stWarning : ST_WARNING_EVENT; // Последнее предупреждение магазина
END_STRUCT
END_TYPE

// Device/Application/ST/ST_HMI/E_HMI_MANUAL_REJECT
{attribute 'qualified_only'}
{attribute 'strict'}
TYPE E_HMI_MANUAL_REJECT :
(
	NONE,
	HMI_OFFLINE,
	MANUAL_MODE_REQUIRED,
	MODBUS_ACTIVE,
	GLOBAL_ERROR_JOG_ONLY,
	DRIVE_ERROR,
	DRIVES_DISABLED,
	AXIS_BUSY,
	AXIS_NOT_HOMED,
	SOFT_LIMIT,
	COMMAND_CONFLICT,
	ROBOT_BUSY,
	ACTION_ALREADY_REACHED,
	EXTERNAL_ROBOT_NOT_READY,
	MOTION_NOT_READY,
	HATCH_CLOSED
);
END_TYPE

// Device/Application/ST/ST_MACHINE/E_MACHINE_OPERATION
{attribute 'qualified_only'}
{attribute 'strict'}
TYPE E_MACHINE_OPERATION :
(
	NONE,
    LOAD,
    UNLOAD,
    CHANGE 
);
END_TYPE

// Device/Application/ST/ST_AXIS/ST_AXIS_FAULT_REQUEST
TYPE ST_AXIS_FAULT_REQUEST :
STRUCT
	xEnabled     : BOOL; // Глобальное разрешение диагностической инъекции
	xJogConflict : BOOL; // Импульс одновременного запроса Jog+ и Jog-
END_STRUCT
END_TYPE

// Device/Application/ST/ST_AXIS_GROUP/ST_AXIS_GROUP_COMMANDS
TYPE ST_AXIS_GROUP_COMMANDS :
STRUCT
	xGlobalError : BOOL; // Глобальная ошибка ячейки
	xPowerPermit : BOOL; // Разрешение включения группы при готовых физических осях
	xEnable      : BOOL; // Импульс включения группы
	xPowerEnable : BOOL; // Импульс включения группы после включения осей FB_AXIS
	xDisable     : BOOL; // Импульс отключения группы
	xReset       : BOOL; // Сброс ошибок группы
	xMoveDirect  : BOOL; // Команда прямого перемещения группы
	xMoveLinear  : BOOL; // Команда линейного перемещения группы
	xHaltCmd     : BOOL; // Команда плавной остановки
	xStopCmd     : BOOL; // Команда остановки группы
END_STRUCT
END_TYPE

// Device/Application/ST/ST_MAGAZINE/ST_TWO_PALLET_COMMAND
TYPE ST_TWO_PALLET_COMMAND :
STRUCT
	xEnable : BOOL;
	xConfirm : BOOL;
	xStart : BOOL; // Атомарно подтвердить актуальную расстановку и включить магазин
	xRejectStart : BOOL; // Оператор ответил «Нет» в предпусковом окне
	xDisable : BOOL;
	xSwap : BOOL;
	xPowerOn : BOOL;
	xPowerOff : BOOL;
	xDriveReset : BOOL;
	xHome : BOOL;
	xLower : BOOL;
	xRaise : BOOL;
	xSelectPallet : BOOL;
	xLockIn : BOOL;
	xLockOut : BOOL;
	xStopIn : BOOL;
	xStopOut : BOOL;
	xMoveToExchange : BOOL;
	xMoveToWork : BOOL;
	xStop : BOOL;
	xReset : BOOL;
	xJogPositive : BOOL;
	xJogNegative : BOOL;
	xJogRelease : BOOL;
	xTeachOperator : BOOL; // Запомнить текущую координату переключения/операторской зоны
	xTeachWork : BOOL; // Запомнить текущую рабочую координату выбранной палеты у робота
	uiPallet : UINT; // Номер подтверждаемой/выбираемой палеты, 1..2
	udiRevision : UDINT; // Ревизия расстановки для команды подтверждения
END_STRUCT
END_TYPE

// Device/Application/ST/ST_MULTI_TYPE/ST_MULTI_TYPE_COMMAND
TYPE ST_MULTI_TYPE_COMMAND :
STRUCT
	{attribute 'symbol' := 'read'}
	xSetTypeCount         : BOOL; // Импульс изменения количества типов
	uiRequestedTypeCount : UINT; // Требуемое количество типов, 1..3
	{attribute 'symbol' := 'read'}
	xSetMachineType       : BOOL; // Импульс назначения типа станку
	uiRequestedMachine   : UINT; // Номер редактируемого станка, 1..3
	uiRequestedMachineType : UINT; // Тип, назначаемый станку
	{attribute 'symbol' := 'read'}
	xSetSlotType          : BOOL; // Импульс назначения типа слоту
	uiRequestedSlot      : UINT; // Номер редактируемого слота
	uiRequestedSlotType  : UINT; // Тип, назначаемый слоту
	{attribute 'symbol' := 'read'}
	xAutoDistribute      : BOOL; // Импульс распределения слотов пропорционально станкам
END_STRUCT
END_TYPE

// Device/Application/ST/ST_AXIS_GROUP/ST_AXIS_GROUP
TYPE ST_AXIS_GROUP :
STRUCT
	Command     : ST_AXIS_GROUP_COMMANDS; // Команды группы осей
	Status      : ST_AXIS_GROUP_STATUS; // Рабочие статусы группы
	Diag        : ST_AXIS_GROUP_DIAGNOSTICS; // Состояние автомата и диагностика
	Error       : ST_AXIS_GROUP_ERRORS; // Активные и последние ошибки
	MotionParam : ST_AXIS_GROUP_MOTION_PARAMS; // Параметры движения
	Timeouts    : ST_AXIS_GROUP_TIMEOUTS; // Допустимое время выполнения шагов
END_STRUCT
END_TYPE

// Device/Application/ST/ST_MAGAZINE/ST_MAGAZINE_FAULT_REQUEST
TYPE ST_MAGAZINE_FAULT_REQUEST :
STRUCT
	xEnabled        : BOOL; // Глобальное разрешение диагностической инъекции
	xWrongOperation : BOOL; // Импульс недопустимой операции
	xNoBlank        : BOOL; // Импульс отсутствия заготовки
	xNoFreeSlot     : BOOL; // Импульс отсутствия свободного слота
	xInvalidSlot    : BOOL; // Импульс недопустимого номера слота
	xSlotContent    : BOOL; // Импульс несоответствия содержимого слота
	xGeometry       : BOOL; // Импульс недопустимой геометрии магазина
END_STRUCT
END_TYPE

// Device/Application/ST/ST_GEOMETRY_CONTROL/ST_GEOMETRY_MEMORY
TYPE ST_GEOMETRY_MEMORY :
STRUCT
	xOccupied : BOOL;
	xRecoveryRequired : BOOL;
	xAtEndSeen : BOOL; // Потерю датчика считаем изъятием только после прихода на него
	dwAlarm : DWORD;
	xRobotStopLatched : BOOL;
	udiLastDepositId : UDINT;
	udiProducedPartsTotal : UDINT;
	Part : ST_GEOMETRY_CALL;
END_STRUCT
END_TYPE

// Device/Application/ST/ST_POINT_MANAGER/E_POINT_MANAGER_STATE
{attribute 'qualified_only'}
{attribute 'strict'}
TYPE E_POINT_MANAGER_STATE :
(
	IDLE,
	SELECT_POINT,
	CHECK_VEL_FACTOR,
	CHECK_ZONE,
	CHECK_ALL
);
END_TYPE

// Device/Application/ST/ST_ALARM/E_ALARM_SEVERITY
TYPE E_ALARM_SEVERITY :
(
	ALARM, // Авария, требующая устранения причины
	WARNING // Предупреждение оператору
);
END_TYPE

// Device/Application/ST/ST_GEOMETRY_CONTROL/ST_GEOMETRY_STATUS
TYPE ST_GEOMETRY_STATUS :
STRUCT
	uiState : UINT; // 0 выключен, 1 свободен, 2 передача роботом, 3 транспорт, 4 ждёт изъятия, 5 восстановление, 6 авария, 7 ручной ход
	xEnabled : BOOL;
	xReady : BOOL;
	xOccupied : BOOL;
	xPartStored : BOOL; // Подтверждённая укладка, отдельно от резерва и неизвестности
	xReserved : BOOL;
	xPartAtEnd : BOOL;
	xDriveRunning : BOOL;
	xDriveAlarm : BOOL;
	xError : BOOL;
	xRobotStopRequired : BOOL;
	xEnableAllowed : BOOL;
	xDisableAllowed : BOOL;
	xConfirmAllowed : BOOL;
	xConfirmationActive : BOOL;
	xRecoveryRequired : BOOL; // Проверка всей ленты нужна независимо от попытки включения
	xManualStartAllowed : BOOL;
	xResetAllowed : BOOL;
	xResetBusy : BOOL;
	xConfigAllowed : BOOL;
	xPointWriteAllowed : BOOL; // Запись данных: связь/SoftMotion/валидные лимиты, без технологических блокировок
	xSimulationRemoveAllowed : BOOL;
	xSimulationAlarmAllowed : BOOL;
	xConfigured : BOOL;
	udiProducedPartsTotal : UDINT;
	udiPartId : UDINT;
	uiMachine : UINT;
	uiProductType : UINT;
	rTravel : REAL; // Положение модели 0..1; в NORMAL только оценка для изображения
	dwEnableBlockers : DWORD; // Причины запрета команды включения; 0 = xEnableAllowed
	dwConfirmBlockers : DWORD; // Причины запрета подтверждения пустоты; 0 = xConfirmAllowed
	xCallWaitWarning : BOOL; // Активный W52 ячейки; снимается подтверждением предупреждений
END_STRUCT
END_TYPE

// Device/Application/ST/ST_STATISTIC/ST_STATISTIC_MACHINE
TYPE ST_STATISTIC_MACHINE :
STRUCT
	rLoadCNC_1            : REAL; // Процент загрузки станка 1
	rLoadCNC_2            : REAL; // Процент загрузки станка 2
	rLoadCNC_3            : REAL; // Процент загрузки станка 3
END_STRUCT
END_TYPE

// Device/Application/ST/ST_MACHINE/ST_MACHINE_SIM_DIAG
TYPE ST_MACHINE_SIM_DIAG :
STRUCT
	xDoorOpening   : BOOL; // Выполняется открытие роботного люка
	xDoorClosing   : BOOL; // Выполняется закрытие роботного люка
	xSafetyDoorOpening : BOOL; // Выполняется открытие операторской двери
	xSafetyDoorClosing : BOOL; // Выполняется закрытие операторской двери
	xChuckClamping : BOOL; // Выполняется зажим патрона
	xChuckOpening  : BOOL; // Выполняется разжим патрона
	xCycleStarting : BOOL; // Выполняется запуск цикла
	xResetAllowed  : BOOL; // Источник имитации снят и авария симулятора может быть сброшена
END_STRUCT
END_TYPE

// Device/Application/ST/ST_MAGAZINE/ST_DETAIL/E_DETAIL_TYPE
{attribute 'qualified_only'}
{attribute 'strict'}
TYPE E_DETAIL_TYPE :
(
	NONE,
	BLANK,
	DETAIL
);
END_TYPE

// Device/Application/ST/ST_GEOMETRY_CONTROL/ST_GEOMETRY_CONFIG
TYPE ST_GEOMETRY_CONFIG :
STRUCT
	xConfigured : BOOL;
	lrX : LREAL;
	lrY : LREAL;
	lrZ : LREAL;
	lrSafeZ : LREAL := -300.0; // Signed-смещение безопасного подхода от рабочей Z
	lrChangeZ : LREAL := -150.0; // Legacy-поле OPC UA; маршрут использует SAFE_Z, при записи равно lrSafeZ
	lrSpeedFactor : LREAL := 0.2;
END_STRUCT
END_TYPE

// Device/Application/ST/ST_AXIS_GROUP/ST_AXIS_GROUP_TIMEOUTS
TYPE ST_AXIS_GROUP_TIMEOUTS :
STRUCT
    tPowerTimeout : TIME := T#5S; // Время ожидания включения или отключения питания
	tGroupTimeout : TIME := T#5S; // Время ожидания включения или отключения группы
    tStopTimeout  : TIME := T#5S; // Время ожидания остановки
	tHaltTimeout  : TIME := T#5S; // Время ожидания плавной остановки
    tHomeTimeout  : TIME := T#30S; // Время ожидания поиска домашней позиции
    tMoveTimeout  : TIME := T#30S; // Время ожидания завершения перемещения
END_STRUCT
END_TYPE

// Device/Application/ST/ST_AXIS_GROUP/ST_AXIS_GROUP_FAULT_REQUEST
TYPE ST_AXIS_GROUP_FAULT_REQUEST :
STRUCT
	xEnabled : BOOL; // Глобальное разрешение диагностической инъекции
	xExecute : BOOL; // Импульс формирования тестовой ошибки SM3
END_STRUCT
END_TYPE

// Device/Application/ST/ST_POINT_MANAGER/ST_POINT_MANAGER_ERRORS
TYPE ST_POINT_MANAGER_ERRORS :
STRUCT
	dwErrorActive : DWORD; // Битовая маска активных ошибок
	dwErrorLast   : DWORD; // Битовая маска последних ошибок
	dwAlarmActive : DWORD; // Собственные аварии менеджера точек для общего журнала
	stErrorActive : ST_POINT_MANAGER_ERROR; // Расшифровка активных ошибок
	stErrorLast   : ST_POINT_MANAGER_ERROR; // Расшифровка последних ошибок
END_STRUCT
END_TYPE

// Device/Application/ST/ST_MACHINE/ST_MACHINE_ERROR
TYPE ST_MACHINE_ERROR :
STRUCT
	WRONG_OPERATION : BOOL; // Не удалось выбрать операцию
	WRONG_COMMAND   : BOOL; // В рецепте встретилась неизвестная команда
	ROBOT_MOTION    : BOOL; // Ошибка перемещения робота
	ROBOT_ACTION    : BOOL; // Ошибка действия захвата
	DOOR_OPEN       : BOOL; // Не удалось открыть дверь
	DOOR_CLOSE      : BOOL; // Не удалось закрыть дверь
	CHUCK_OPEN      : BOOL; // Не удалось разжать патрон
	CHUCK_CLOSE     : BOOL; // Не удалось зажать патрон
	CYCLE_START     : BOOL; // Не удалось запустить цикл станка
	SAFETY_STOP     : BOOL; // Получена глобальная ошибка ячейки
	UNKNOWN_DETAIL  : BOOL; // Неизвестно состояние детали в станке
	MACHINE_ALARM   : BOOL; // Станок сообщил аварию
	INDEX_ERROR     : BOOL; // Индекс рецепта вышел за границы
	DOOR_ROBOT      : BOOL; // Дверь закрыта при нахождении робота внутри
	MACHINE_IDLE    : BOOL; // Авария станка возникла в ожидании
	TIMEOUT_ROBOT_MOVE    : BOOL; // Превышено время перемещения робота
	TIMEOUT_ROBOT_ACTION  : BOOL; // Превышено время действия захвата
	TIMEOUT_ROBOT_RELEASE : BOOL; // Робот не освободил интерфейс команды вовремя
	TIMEOUT_DOOR_OPEN     : BOOL; // Превышено время открытия двери
	TIMEOUT_DOOR_CLOSE    : BOOL; // Превышено время закрытия двери
	TIMEOUT_HATCH_UNLOCK  : BOOL; // Превышено время открытия замка роботного люка
	TIMEOUT_CHUCK_OPEN    : BOOL; // Превышено время разжима патрона
	TIMEOUT_CHUCK_CLOSE   : BOOL; // Превышено время зажима патрона
	TIMEOUT_CYCLE_START   : BOOL; // Превышено время подтверждения запуска цикла
	SAFETY_DOOR_OPEN     : BOOL; // Операторская дверь открылась во время обслуживания
	HATCH_UNLOCK_PROCESSING : BOOL; // Замок открыт во время обработки в автоматической линии
END_STRUCT
END_TYPE

// Device/Application/ST/ST_AXIS_GROUP/ST_AXIS_GROUP_MOTION_PARAMS
TYPE ST_AXIS_GROUP_MOTION_PARAMS :
STRUCT
	stTargetPos      : SMC_POS_REF; // Целевая позиция в формате SoftMotion
	lrX              : LREAL := 1000; // Целевая координата X
	lrY              : LREAL := 1000; // Целевая координата Y
	lrZ              : LREAL := 1000; // Целевая координата Z
	VelFactor        : LREAL := 0.1; // Коэффициент скорости
	AccFactor        : LREAL := 0.1; // Коэффициент ускорения
	JerkFactor       : LREAL := 0.1; // Коэффициент рывка
	HaltDeceleration : LREAL := 1000; // Замедление при плавной остановке
	HaltJerk         : LREAL := 10000; // Рывок при плавной остановке
END_STRUCT
END_TYPE

// Device/Application/ST/ST_TEST/ST_TEST_SCENARIO_BUFFER
TYPE ST_TEST_SCENARIO_BUFFER :
STRUCT
	udiLoadSeq : UDINT;
	uiTypeCount : UINT;
	axMagazineEnabled : ARRAY [1..2] OF BOOL;
	auiMachineState : ARRAY [1..3] OF UINT; // 0 disabled, 1 empty, 2 blank processing, 3 detail ready
	auiMachineType : ARRAY [1..3] OF UINT;
	aauiSlotContent : ARRAY [1..2, 1..120] OF UINT; // Две статичные кассеты: 0 empty, 1 blank, 2 detail
	auiSlotType : ARRAY [1..120] OF UINT;
	auiGripperContent : ARRAY [1..2] OF UINT;
	auiGripperType : ARRAY [1..2] OF UINT;
	uiOrientation : UINT; // 0 blank, 1 detail
	dwCellFaultMask : DWORD; // b0: противоречивое наличие детали в обоих захватах
	dwRobotFaultMask : DWORD; // b0 wrong action; b1..b4 grippers; b5..b8 point validation
	adwMagazineFaultMask : ARRAY [1..2] OF DWORD; // b0 wrong op; b1 no blank; b2 no slot; b3 invalid slot; b4 content; b5 geometry
	adwMachineFaultMask : ARRAY [1..3] OF DWORD; // b0 alarm; b1 door; b2 chuck; b3..b10 timeouts
END_STRUCT
END_TYPE

// Device/Application/ST/ST_CELL/ST_CONTROL_CABINET_IO_STATUS
TYPE ST_CONTROL_CABINET_IO_STATUS :
STRUCT
	xEmergencyStopPressed : BOOL; // Нормализованный вход: TRUE — грибок нажат
	xStartPressed         : BOOL; // Физическая кнопка «Включить ячейку»
	xStopPressed          : BOOL; // Физическая кнопка «Выключить ячейку»
	xResetPressed         : BOOL; // Физическая кнопка общего сброса ошибок
END_STRUCT
END_TYPE

// Device/Application/ST/ST_MAGAZINE/ST_TWO_PALLET_DIAG
TYPE ST_TWO_PALLET_DIAG :
STRUCT
	eState : E_TWO_PALLET_STATE := E_TWO_PALLET_STATE.IDLE;
	eFaultState : E_TWO_PALLET_STATE := E_TWO_PALLET_STATE.IDLE;
	uiReason : UINT; // Первая причина блокировки подтверждения/включения магазина
	stWarning : ST_WARNING_EVENT;
END_STRUCT
END_TYPE

// Device/Application/ST/ST_CELL/ST_CELL_STATUS
TYPE ST_CELL_STATUS :
STRUCT
	xMagazineExchangeAllowed : BOOL; // Планировщик не держит незавершённый маршрут
	xRunning           : BOOL; // Автоматический цикл запущен
	xStopPending       : BOOL; // Запрошена остановка после безопасного шага
	xBusy              : BOOL; // Менеджер выполняет автоматический цикл
	xWaitingMachine    : BOOL; // Ожидание доступного станка
	xWaitingMagazine   : BOOL; // Ожидание пополнения или освобождения магазина
	xError             : BOOL; // Менеджер ячейки находится в ошибке
	xReadyToStart      : BOOL; // Выполнены все условия запуска автоматического цикла
	xStartAllowed      : BOOL; // Кнопка запуска или отмены ожидающей остановки доступна
	xStopAllowed       : BOOL; // Кнопка остановки автоматического цикла доступна
	xResetAllowed      : BOOL; // Кнопка общего сброса доступна
	xManualAllowed     : BOOL; // Кнопка перехода в ручной режим доступна
	xAutomaticAllowed  : BOOL; // Кнопка перехода в автоматический режим доступна
	xDrivesReady       : BOOL; // Приводы и группа осей готовы к движению
	xRobotReady        : BOOL; // Робот готов принять команду
	xMagazineReady     : BOOL; // Магазин готов к работе с роботом
	xSafetyHomeRequired: BOOL; // Повторный запуск разрешён только из HOME_SAFETY
	xRobotAtSafetyHome : BOOL; // Фактические координаты находятся в диапазоне HOME_SAFETY
	xStartCheckCellIdle          : BOOL; // Менеджер ячейки готов принять новый запуск
	xStartCheckAutomaticMode     : BOOL; // Выбран автоматический режим
	xStartCheckNoBlockingError   : BOOL; // Нет блокирующей запуск ошибки
	xStartCheckRobotInterfaceReady: BOOL; // Выбранный интерфейс робота готов
	xStartCheckConfigurationValid: BOOL; // Конфигурация типов корректна
	xStartCheckPointsConfigured  : BOOL; // HOME_SAFETY и точки включённого оборудования настроены
	xStartCheckDrivesReady       : BOOL; // Приводы и группа готовы
	xStartCheckRobotReady        : BOOL; // Робот готов принять маршрут
	xStartCheckMagazineReady     : BOOL; // Магазин готов к операции
	xStartCheckTaskAvailable     : BOOL; // Есть допустимая работа или известный груз
	xStartCheckSafetyHome        : BOOL; // Условие HOME_SAFETY выполнено
	xStartCheckSafety            : BOOL; // Грибки, реле и двери безопасности готовы
	uiStartConditionsMet        : UINT; // Количество выполненных условий запуска
	uiStartConditionsTotal      : UINT; // Общее количество условий запуска
	uiReadyMachines    : UINT; // Количество включённых станков в состоянии IDLE
	uiSelectedMachine  : UINT; // Номер выбранного станка
	uiActiveMagazine   : UINT; // Магазин, закреплённый за текущим автоматическим циклом
	eMagazineOperation : E_MAGAZINE_OPERATION; // Выбранная операция магазина
	xOperatorPromptActive : BOOL; // PLC ожидает ответ оператора перед запуском цикла
	xOperatorChoiceAllowed: BOOL; // PLC разрешает отправить вариант активного опроса
	xOperatorCancelAllowed: BOOL; // PLC разрешает отменить активный предпусковой опрос
	uiOperatorPrompt      : UINT; // 0 нет; 1/3 содержимое захвата; 2/4 тип; 5 станок
	uiOperatorTypeMask    : UINT; // Биты 0..2 — доступные типы продукции
	uiOperatorMachineMask : UINT; // Биты 0..2 — допустимые станки для стартового LOAD
END_STRUCT
END_TYPE

// Device/Application/ST/ST_ROBOT/E_ROBOT_STATE
{attribute 'qualified_only'}
{attribute 'strict'}
TYPE E_ROBOT_STATE :
(
	IDLE,
	MOTION,
	GRIPPER,
	DONE,
    ERROR,
	MODBUS
);
END_TYPE

// Device/Application/ST/ST_MULTI_TYPE/ST_MULTI_TYPE_CONFIG
TYPE ST_MULTI_TYPE_CONFIG :
STRUCT
	uiTypeCount    : UINT; // Количество типов обрабатываемых деталей, 1..3
	auiMachineType : ARRAY [1..3] OF UINT; // Тип, закреплённый за каждым станком
	auiSlotType    : ARRAY [1..GVL_CELL_SETTINGS.NumberDetail] OF UINT; // Тип заготовки каждого слота
END_STRUCT
END_TYPE

// Device/Application/ST/ST_MACHINE/ST_MACHINE_RECIPE
TYPE ST_MACHINE_RECIPE :
STRUCT
	eRobotAction    : E_ROBOT_ACTION; // Действие робота на шаге рецепта
	eCommand        : E_MACHINE_STATE; // Команда шага рецепта
	stPoint         : E_MACHINE_POINTS; // Логическая точка станка
	xRetreatStarted : BOOL; // Признак начала отхода робота
	xRobotDone      : BOOL; // Признак освобождения робота после шага
END_STRUCT
END_TYPE

// Device/Application/ST/ST_AXIS/ST_AXIS
TYPE ST_AXIS :
STRUCT
	Command     : ST_AXIS_COMMANDS; // Команды оси
	Status      : ST_AXIS_STATUS; // Рабочие статусы оси
	Diag        : ST_AXIS_DIAGNOSTICS; // Состояние автомата и текстовая диагностика
	Error       : ST_AXIS_ERROR_CODES; // Активные и последние ошибки
	MotionParam : ST_AXIS_MOTION_PARAMS; // Параметры движения
	Timeouts    : ST_AXIS_TIMEOUTS; // Допустимое время выполнения шагов

END_STRUCT
END_TYPE

// Device/Application/ST/ST_POINT_MANAGER/ST_POINT_MANAGER
TYPE ST_POINT_MANAGER :
STRUCT
	Command : ST_POINT_MANAGER_COMMAND; // Команды менеджера точки
	Status  : ST_POINT_MANAGER_STATUS; // Рабочие статусы менеджера точки
	Diag    : ST_POINT_MANAGER_DIAG; // Состояние автомата и допустимые пределы
	Error   : ST_POINT_MANAGER_ERRORS; // Активные и последние ошибки
END_STRUCT
END_TYPE

// Device/Application/ST/ST_STATISTIC/ST_STATISTIC_ROBOT
TYPE ST_STATISTIC_ROBOT :
STRUCT
	tCNC_1      	: TIME; // Среднее время работы в стнке 1
	tCNC_2      	: TIME; // Среднее время работы в стнке 2
	tCNC_3      	: TIME; // Среднее время работы в стнке 3
	tMoveCNC_1 		: TIME; // Среднее время перемещения от магазина к станку 1
	tMoveCNC_2 		: TIME; // Среднее время перемещения от магазина к станку 2
	tMoveCNC_3 		: TIME; // Среднее время перемещения от магазина к станку 3
	tMagazine       : TIME; // Среднее время работы в магазине

	rRobot          : REAL; // Процент загрузки робота
END_STRUCT
END_TYPE

// Device/Application/ST/ST_AXIS_GROUP/E_AXIS_GROUP_POWER_MODE
{attribute 'qualified_only'}
{attribute 'strict'}
TYPE E_AXIS_GROUP_POWER_MODE :
(
	OFF,
	OFF_REQUEST,
	ON
	
);
END_TYPE

// Device/Application/ST/ST_POINT/ST_POINT
TYPE ST_POINT :
STRUCT
	Name        : STRING[80]; // Имя точки
	X           : LREAL; // Координата X
	Y           : LREAL; // Координата Y
	Z           : LREAL; // Координата Z
	MagazineSafeZ : LREAL; // Signed-смещение Safe Z базы магазина или ГК
	MagazineChangeZ : LREAL; // Signed-смещение Change Z; используется только базовой точкой магазина
	SpeedFactor : LREAL; // Коэффициент скорости движения
	xConfigured : BOOL; // Для базы магазина TRUE только при ненулевых MagazineSafeZ и MagazineChangeZ
END_STRUCT
END_TYPE

// Device/Application/ST/ST_MAGAZINE/ST_MAGAZINE_ERRORS
TYPE ST_MAGAZINE_ERRORS :
STRUCT
	dwErrorActive : DWORD; // Битовая маска активных ошибок
	dwErrorLast   : DWORD; // Битовая маска последних ошибок
	dwAlarmActive : DWORD; // Собственные аварии магазина для общего журнала
	stErrorActive : ST_MAGAZINE_ERROR; // Расшифровка активных ошибок
	stErrorLast   : ST_MAGAZINE_ERROR; // Расшифровка последних ошибок
END_STRUCT
END_TYPE

// Device/Application/ST/ST_ALARM/ST_WARNING_EVENT
TYPE ST_WARNING_EVENT :
STRUCT
	udiSequence : UDINT; // Порядковый номер предупреждения от функционального блока
	uiCode      : UINT; // Код предупреждения внутри функционального блока
END_STRUCT
END_TYPE

// Device/Application/ST/ST_MULTI_TYPE/ST_MULTI_TYPE_HMI
TYPE ST_MULTI_TYPE_HMI :
STRUCT
	Command      : ST_MULTI_TYPE_COMMAND; // Команды конфигурации от HMI
	Config       : ST_MULTI_TYPE_CONFIG; // Фактически принятая конфигурация
	ConfigStatus : ST_MULTI_TYPE_CONFIG_STATUS; // Разрешения и диагностика конфигурации
	CycleStatus  : ST_CELL_CYCLE_STATUS; // Диагностика универсального цикла
END_STRUCT
END_TYPE

// Device/Application/ST/ST_MACHINE/ST_MACHINE_TIMEOUTS
TYPE ST_MACHINE_TIMEOUTS :
STRUCT
	tRobotMove    : TIME := T#60S; // Допустимое время движения робота
	tRobotAction  : TIME := T#10S; // Допустимое время действия захвата
	tRobotRelease : TIME := T#5S; // Допустимое время освобождения интерфейса робота
	tDoorOpen     : TIME := T#10S; // Допустимое время открытия двери
	tDoorClose    : TIME := T#10S; // Допустимое время закрытия двери
	tHatchUnlock  : TIME := T#5S; // Допустимое ожидание открытия замка роботного люка
	tChuckOpen    : TIME := T#10S; // Допустимое время разжима патрона
	tChuckClose   : TIME := T#10S; // Допустимое время зажима патрона
	tCycleStart   : TIME := T#10S; // Допустимое время подтверждения запуска цикла
END_STRUCT
END_TYPE

// Device/Application/ST/ST_GRIPPER/ST_GRIPPER_FAULT_REQUEST
TYPE ST_GRIPPER_FAULT_REQUEST :
STRUCT
	xEnabled        : BOOL; // Глобальное разрешение диагностической инъекции
	xGripper1Fault  : BOOL; // Неисправность первого захвата
	xGripper2Fault  : BOOL; // Неисправность второго захвата
	xRotationFault  : BOOL; // Неисправность механизма поворота
	xGlobalFault    : BOOL; // Общая неисправность захвата
END_STRUCT
END_TYPE

// Device/Application/ST/ST_HMI/ST_AXIS_HMI_STATUS
TYPE ST_AXIS_HMI_STATUS :
STRUCT
	xJogPositiveAllowed   : BOOL; // PLC разрешает положительный Jog
	xJogNegativeAllowed   : BOOL; // PLC разрешает отрицательный Jog
	xHomeAllowed          : BOOL; // PLC разрешает поиск домашней позиции
	xMoveAbsoluteAllowed  : BOOL; // PLC разрешает абсолютное движение
	xMoveRelativePositiveAllowed : BOOL; // PLC разрешает положительный короткий шаг
	xMoveRelativeNegativeAllowed : BOOL; // PLC разрешает отрицательный короткий шаг
	xDriveReady           : BOOL; // Ось включена и готова к движению
	xBusy                 : BOOL; // Ось выполняет ручную команду
	xError                : BOOL; // На оси есть ошибка
	xHomed                : BOOL; // Ось прошла поиск домашней позиции
	lrActualPosition      : LREAL; // Фактическая координата
	lrTargetPosition      : LREAL; // Принятая целевая координата
	lrDeviation           : LREAL; // Отклонение фактической координаты от цели
	lrMinPosition         : LREAL; // Нижний программный предел
	lrMaxPosition         : LREAL; // Верхний программный предел
	lrCommandVelocity     : LREAL; // Фактически заданная скорость ручного движения
	lrMaxVelocity         : LREAL; // Скорость, соответствующая 100 процентам
	eRejectReason         : E_HMI_MANUAL_REJECT; // Числовая причина недоступности команды
	eState                : E_AXIS_STATE; // Числовое состояние автомата оси
END_STRUCT
END_TYPE

// Device/Application/ST/ST_ALARM/ST_ALARM_SOURCE_DATA
TYPE ST_ALARM_SOURCE_DATA :
STRUCT
	eSource       : E_ALARM_SOURCE; // Функциональный блок, которому принадлежит событие
	dwAlarmActive : DWORD; // Только собственные активные аварии блока
	xRobotStopRequired : BOOL; // Владелец зафиксировал зависимый останов робота для этого контекста
	xGlobalError  : BOOL; // Глобальная ошибка была активна в момент публикации источника
	stWarning     : ST_WARNING_EVENT; // Последнее предупреждение блока
END_STRUCT
END_TYPE

// Device/Application/ST/ST_MAGAZINE/ST_MAGAZINE_COMMAND
TYPE ST_MAGAZINE_COMMAND :
STRUCT
	xEnable  : BOOL; // Импульс включения магазина
	xDisable : BOOL; // Импульс отключения магазина
	xExecute : BOOL; // Запуск выбранной операции
	xStop    : BOOL; // Остановка текущей операции
	eOperation : E_MAGAZINE_OPERATION; // Операция автоматического цикла
	iTakeSlot  : SINT; // Слот заготовки для TAKE/CHANGE
	iPutSlot   : SINT; // Слот укладки для PUT/CHANGE/RETURN_BLANK
END_STRUCT
END_TYPE

// Device/Application/ST/ST_MACHINE/E_MACHINE_STATE
{attribute 'qualified_only'}
{attribute 'strict'}
TYPE E_MACHINE_STATE :
(
	DISABLED := 0,
	OPERATOR_CHOICE_PART,
	OPERATOR_CHOICE_RUN,
	OPERATOR_CHOICE_DOOR,
    IDLE,
	CHOSE,
	READ,
	NEXT,
	RELEASE_ROBOT_ACTION,
	ROBOT_MOVE,
	ROBOT_ACTION,
	DOOR_OPEN,
	DOOR_CLOSE,
	CHUCK_OPEN,
	CHUCK_CLOSE,
	CYCLE_START,
	DONE,
	ERROR
);
END_TYPE

// Device/Application/ST/ST_MAGAZINE/ST_DETAIL/ST_DETAIL
TYPE ST_DETAIL :
STRUCT
	eDetailType : E_DETAIL_TYPE; // Тип содержимого слота
	xInPosition : BOOL; // Признак наличия объекта в слоте
	uiProductType : UINT; // Тип продукции перемещается между зонами вместе со слотом
END_STRUCT
END_TYPE

// Device/Application/ST/ST_TEST/E_CELL_TEST_ENVIRONMENT
{attribute 'qualified_only'}
TYPE E_CELL_TEST_ENVIRONMENT :
(
	NORMAL := 0,
	SIMULATION := 1,
	SC500_BENCH := 2
);
END_TYPE

// Device/Application/ST/ST_GRIPPER/ST_GRIPPER_ERRORS
TYPE ST_GRIPPER_ERRORS :
STRUCT
	dwErrorActive : DWORD; // Битовая маска активных ошибок
	dwErrorLast   : DWORD; // Битовая маска последних ошибок
	dwAlarmActive : DWORD; // Собственные аварии захвата для общего журнала
	stErrorActive : ST_GRIPPER_ERROR; // Расшифровка активных ошибок
	stErrorLast   : ST_GRIPPER_ERROR; // Расшифровка последних ошибок
END_STRUCT
END_TYPE

// Device/Application/ST/ST_AXIS_GROUP/E_AXIS_GROUP_STATE
{attribute 'qualified_only'}
{attribute 'strict'}
TYPE E_AXIS_GROUP_STATE :
(
	DISABLED,
	DISABLING_GROUP,
	DISABLING_POWER,
	ENABLING_POWER,
	ENABLING_GROUP,
	READY,
	MOVING_DIRECT,
	MOVING_LINEAR,
	EMG_STOP,
	HALT_STOP,
	WAIT_STOP,	
	ERROR,
	RESETTING,
	RESET_VERIFY

	
);
END_TYPE

// Device/Application/ST/ST_POINT_MANAGER/ST_POINT_MANAGER_ERROR
TYPE ST_POINT_MANAGER_ERROR :
STRUCT
	X_OUT_OF_LIMIT : BOOL; // Координата X находится вне допустимой зоны
	Y_OUT_OF_LIMIT : BOOL; // Координата Y находится вне допустимой зоны
	Z_OUT_OF_LIMIT : BOOL; // Координата Z находится вне допустимой зоны
	INVALID_VEL    : BOOL; // Коэффициент скорости задан неверно
	X_LIMIT_CONFIG_INVALID : BOOL; // Software limits оси X отключены или заданы некорректно
	Y_LIMIT_CONFIG_INVALID : BOOL; // Software limits оси Y отключены или заданы некорректно
	Z_LIMIT_CONFIG_INVALID : BOOL; // Software limits оси Z отключены или заданы некорректно
	POINT_NOT_CONFIGURED : BOOL; // Инженерная точка ещё не сохранена редактором
END_STRUCT
END_TYPE

// Device/Application/ST/ST_MAGAZINE/E_MAGAZINE_STATE
{attribute 'qualified_only'}
{attribute 'strict'}
TYPE E_MAGAZINE_STATE :
(
	DISABLED,
	IDLE,
	CHOOSE,
	PREPARE_STEP,
	ROBOT_COMMAND,
	RELEASE_ROBOT_COMMAND,
	NEXT,
	DONE,
	ERROR
);
END_TYPE

// Device/Application/ST/ST_GEOMETRY_CONTROL/ST_GEOMETRY_SIGNALS
TYPE ST_GEOMETRY_SIGNALS :
STRUCT
	xReserve : BOOL;
	xDeposited : BOOL;
	xReleased : BOOL;
	xRobotInteraction : BOOL;
	Call : ST_GEOMETRY_CALL;
END_STRUCT
END_TYPE

// Device/Application/ST/ST_ROBOT/ST_ROBOT_COMMAND
TYPE ST_ROBOT_COMMAND :
STRUCT
	xExecute : BOOL; // Команда запуска
	xStop    : BOOL; // Команда остановки
	xReset   : BOOL; // Команда сброса внешнего робота
	eAction  : E_ROBOT_ACTION; // Элементарное действие робота
	eSetPoint: E_POINT_NAME; // Имя элементарной точки движения
	iActiveSlot : SINT; // Единственный слот, относительно которого выполняется команда
	uiMagazineId : UINT; // 0 вне магазина; 1 или 2 для точки соответствующего магазина
END_STRUCT
END_TYPE

// Device/Application/ST/ST_CELL/ST_CELL_SAFETY_STATUS
TYPE ST_CELL_SAFETY_STATUS :
STRUCT
	xReady                   : BOOL; // Все текущие условия безопасности выполнены
	xGlobalError             : BOOL; // Хотя бы одна текущая Safety-причина активна
	xPhaseRelayOk            : BOOL; // Реле контроля фаз в норме
	xPressureRelayOk         : BOOL; // Реле контроля давления в норме
	xSafetyRelayOk           : BOOL; // Реле безопасности взведено
	xSafetyRelayResetAllowed : BOOL; // Разрешён отдельный импульс сброса реле
	xSafetyRelayResetActive  : BOOL; // Полный секундный импульс сброса реле сейчас активен
	axEmergencyStopReleased  : ARRAY [1..7] OF BOOL; // 4 поста, 2 шкафа, MPG
	axDoorReady              : ARRAY [1..4] OF BOOL; // Замок закрыт либо связанный магазин выключен
	axButtonStationPressed   : ARRAY [1..4] OF BOOL; // Фактический вход кнопки поста, с учётом симуляции
	axButtonStationLightOn   : ARRAY [1..4] OF BOOL; // Выход подсветки кнопки поста
END_STRUCT
END_TYPE

// Device/Application/ST/ST_TEST/E_TEST_SPEED_PROFILE
{attribute 'qualified_only'}
TYPE E_TEST_SPEED_PROFILE :
(
	REALTIME := 0,
	FAST := 1
);
END_TYPE

// Device/Application/ST/ST_AXIS_GROUP/ST_AXIS_GROUP_STATUS
TYPE ST_AXIS_GROUP_STATUS :
STRUCT
	xLocalError     : BOOL; // Активна любая внутренняя ошибка блока
	xLogicalError   : BOOL; // Активна логическая ошибка группы
	xGroupError     : BOOL; // Активна ошибка SoftMotion группы
	xMoveDirectDone : BOOL; // Прямое перемещение завершено
	xSimErrorAllowed: BOOL; // Разрешена безопасная тестовая инъекция ошибки SM3
	xPositionValid  : BOOL; // Координаты группы подтверждены MC_GroupReadActualPosition
	ActualX         : LREAL; // Текущая координата X
	ActualY         : LREAL; // Текущая координата Y
	ActualZ         : LREAL; // Текущая координата Z
	
END_STRUCT
END_TYPE

// Device/Application/ST/ST_MACHINE/ST_MACHINE_DIAG
TYPE ST_MACHINE_DIAG :
STRUCT
	eState            : E_MACHINE_STATE; // Текущее состояние автомата станка
	eGrantedOperation : E_MACHINE_OPERATION; // Разрешённая операция
	eActualOperation  : E_MACHINE_OPERATION; // Выполняемая операция
	stWarning         : ST_WARNING_EVENT; // Последнее предупреждение станка
END_STRUCT
END_TYPE

// Device/Application/ST/ST_MACHINE/ST_MACHINE_IO_COMMAND
TYPE ST_MACHINE_IO_COMMAND :
STRUCT
	xOpenDoor       : BOOL; // Открыть роботный люк; имя сохранено для совместимости
	xCloseDoor      : BOOL; // Закрыть роботный люк; имя сохранено для совместимости
	xHatchUnLock    : BOOL; // Открыть замок роботного люка; FALSE удерживает замок закрытым
	xOpenSafetyDoor : BOOL; // Открыть операторскую дверь
	xCloseSafetyDoor: BOOL; // Закрыть операторскую дверь
	xClampChuck   : BOOL; // Зажать патрон
	xUnclampChuck : BOOL; // Разжать патрон
	xStartCycle   : BOOL; // Запустить обработку
	xReset        : BOOL; // Сбросить аварию станка
END_STRUCT
END_TYPE

// Device/Application/ST/ST_AXIS_GROUP/E_MOTION_RESET_STATE
{attribute 'qualified_only'}
{attribute 'strict'}
TYPE E_MOTION_RESET_STATE :
(
	IDLE,
	RESET_GROUP,
	WAIT_GROUP,
	RESET_AXES,
	WAIT_AXES
);
END_TYPE

// Device/Application/ST/ST_ALARM/E_ALARM_SOURCE
TYPE E_ALARM_SOURCE :
(
	CELL, // Ячейка
	ROBOT, // Робот
	MACHINE_1, // Станок 1
	MACHINE_2, // Станок 2
	MACHINE_3, // Станок 3
	MAGAZINE_LOGIC_1, // Магазин 1; имя не конфликтует с SoftMotion-осью Magazine_1
	MAGAZINE_LOGIC_2, // Магазин 2; имя не конфликтует с SoftMotion-осью Magazine_2
	RESERVED_LEGACY_MAGAZINE_AXIS_1, // Код 7 сохранён только для старых записей журнала
	RESERVED_LEGACY_MAGAZINE_AXIS_2, // Код 8 сохранён только для старых записей журнала
	AXIS_X, // Ось X
	AXIS_Y, // Ось Y
	AXIS_Z, // Ось Z
	AXIS_GROUP, // Группа осей XYZ
	MOTION_MANAGER, // Менеджер движения
	POINT_MANAGER, // Менеджер точек
	GRIPPER, // Захват робота
	CELL_SAFETY, // Дискретный контур безопасности; прежние числовые коды сохранены
	GEOMETRY_1,
	GEOMETRY_2
);
END_TYPE

// Device/Application/ST/ST_CELL/ST_MPG_IO_STATUS
TYPE ST_MPG_IO_STATUS :
STRUCT
	xEmergencyStopPressed : BOOL; // Нормализованный вход: TRUE — грибок MPG нажат
	xAxisX                : BOOL; // Положение селектора оси X
	xAxisY                : BOOL; // Положение селектора оси Y
	xAxisZ                : BOOL; // Положение селектора оси Z
	xMultiplier1          : BOOL; // Положение множителя x1
	xMultiplier10         : BOOL; // Положение множителя x10
	xMultiplier100        : BOOL; // Положение множителя x100
END_STRUCT
END_TYPE

// Device/Application/ST/ST_ROBOT/ST_ROBOT_ERROR
TYPE ST_ROBOT_ERROR :
STRUCT
	WRONG_ACTION : BOOL; // Получена неизвестная команда робота
	MOTION_ERROR : BOOL; // Ошибка менеджера движения
	GRIPPER_ERROR: BOOL; // Ошибка механизма захвата
	MODBUS_ERROR : BOOL; // Совместимость: любая ошибка внешнего интерфейса
	MODBUS_COMMUNICATION_ERROR : BOOL; // Ошибка TCP/FC03/FC16/heartbeat
	EXTERNAL_ROBOT_ALARM : BOOL; // Контроллер робота сообщил технологическую аварию
	STOP_ERROR   : BOOL; // Движение остановлено командой или глобальной ошибкой
END_STRUCT
END_TYPE

// Device/Application/ST/ST_MOTION_MANAGER/ST_MOTION_MANAGER_ERRORS
TYPE ST_MOTION_MANAGER_ERRORS :
STRUCT
	dwErrorActive : DWORD; // Битовая маска активных ошибок
	dwErrorLast   : DWORD; // Битовая маска последних ошибок
	dwAlarmActive : DWORD; // Собственные аварии менеджера движения для общего журнала
	stErrorActive : ST_MOTION_MANAGER_ERROR; // Расшифровка активных ошибок
	stErrorLast   : ST_MOTION_MANAGER_ERROR; // Расшифровка последних ошибок
END_STRUCT
END_TYPE

// Device/Application/ST/ST_MACHINE/ST_MACHINE_FAULT_REQUEST
TYPE ST_MACHINE_FAULT_REQUEST :
STRUCT
	xEnabled             : BOOL; // Глобальное разрешение диагностической инъекции
	xReset               : BOOL; // Отдельный сброс источника неисправности станка
	xMachineAlarm        : BOOL; // Общая авария виртуального станка
	xDoorFault           : BOOL; // Неисправность механизма двери
	xChuckFault          : BOOL; // Неисправность механизма патрона
	xTimeoutRobotMove    : BOOL; // Не подтверждать завершение движения робота
	xTimeoutRobotAction  : BOOL; // Не подтверждать действие захвата
	xTimeoutRobotRelease : BOOL; // Не подтверждать освобождение интерфейса робота
	xTimeoutDoorOpen     : BOOL; // Не подтверждать открытие двери
	xTimeoutDoorClose    : BOOL; // Не подтверждать закрытие двери
	xTimeoutHatchUnlock  : BOOL; // Не подтверждать открытие замка до TIMEOUT
	xTimeoutChuckOpen    : BOOL; // Не подтверждать разжим патрона
	xTimeoutChuckClose   : BOOL; // Не подтверждать зажим патрона
	xTimeoutCycleStart   : BOOL; // Не подтверждать запуск цикла обработки
END_STRUCT
END_TYPE

// Device/Application/ST/ST_MAGAZINE/E_TWO_PALLET_STATE
{attribute 'qualified_only'}
{attribute 'strict'}
TYPE E_TWO_PALLET_STATE :
(
	IDLE := 0,
	AUTO_LOWER := 20,
	AUTO_MOVE_TO_EXCHANGE := 30,
	AUTO_SELECT_PALLET := 40,
	AUTO_MOVE_TO_WORK := 50,
	AUTO_RAISE := 60,
	MANUAL_LOWER := 100,
	MANUAL_RAISE := 110,
	MANUAL_SELECT_PALLET := 120,
	MANUAL_MOVE := 130,
	MANUAL_HOME := 150,
	MANUAL_JOG := 160,
	MANUAL_LOCK := 170,
	MANUAL_STOP := 180
);
END_TYPE

// Device/Application/ST/ST_MAGAZINE/ST_TWO_PALLET_CONFIG
TYPE ST_TWO_PALLET_CONFIG :
STRUCT
	xConfigured : BOOL; // Не выставляется автоматически; параметры проверены на механизме
	xP1LockOut : BOOL; // Legacy: используется только при переносе старой RETAIN-конфигурации
	lrExchange : LREAL;
	lrWorkP1 : LREAL;
	lrWorkP2 : LREAL;
	lrHome : LREAL;
	lrTolerance : LREAL;
	lrVelocity : LREAL;
	lrAcceleration : LREAL;
	lrDeceleration : LREAL;
	lrJerk : LREAL;
	tCylinder : TIME;
	tMove : TIME;
	tHome : TIME;
	tPulse : TIME;
	xSignalPatternsConfigured : BOOL;
	uiP1Signals : UINT; // Биты 0..5: LiftDown, LiftUp, LockIn, LockOut, StopIn, StopOut
	uiP2Signals : UINT; // Полные ожидаемые состояния шести герконов для П2 у робота
END_STRUCT
END_TYPE

// Device/Application/ST/ST_ROBOT/E_ROBOT_ACTION
{attribute 'qualified_only'}
{attribute 'strict'}
TYPE E_ROBOT_ACTION :
(
	NONE,
	MOVE_TO_POINT,
	UNCLAMP_1,
	CLAMP_1,
	UNCLAMP_2,
	CLAMP_2,
	ROTATE_TO_BLANK,
	ROTATE_TO_DETAIL
					
);
END_TYPE

// Device/Application/ST/ST_AXIS/ST_AXIS_STATUS
TYPE ST_AXIS_STATUS :
STRUCT
	xStandstill : BOOL; // MC_ReadStatus: подтверждённый останов, включая Disabled/ErrorStop
    xPowered            : BOOL; // На привод подано питание
	xPowerStageOn        : BOOL; // Фактическое подтверждение включения силовой части
	xDriveStartOn        : BOOL; // Фактическое подтверждение снятого QuickStop
	xPowerOff            : BOOL; // Силовая часть отключена и QuickStop активен
    xBusy               : BOOL; // Ось выполняет команду
    xDone               : BOOL; // Последняя команда завершена
    xError              : BOOL; // Активна любая ошибка оси
    xHomed              : BOOL; // Ось прошла поиск домашней позиции
    xLocalError         : BOOL; // Активна внутренняя ошибка блока
    xMotionBusy         : BOOL; // Активен один из блоков движения
    xCanStartMotion     : BOOL; // Разрешён запуск новой команды движения
    xAxisError          : BOOL; // Активна ошибка привода или SoftMotion
    xLogicalError       : BOOL; // Активна логическая ошибка блока
    xWarning            : BOOL; // Активно предупреждение
    xAxisResetNeeded    : BOOL; // Требуется сброс ошибки привода
    xLogicalResetNeeded : BOOL; // Требуется сброс логической ошибки
	lrActualPosition    : REAL; // Текущая позиция оси
END_STRUCT
END_TYPE

// Device/Application/ST/ST_FAULT_INJECTOR/ST_FAULT_INJECTION_STATUS
TYPE ST_FAULT_INJECTION_STATUS :
STRUCT
	xAllowed          : BOOL; // Инъекция разрешена текущим состоянием владельца
	xActive           : BOOL; // Источник тестовой неисправности активен
	xBusy             : BOOL; // Выполняется одноразовый сценарий инъекции
	xResetAllowed     : BOOL; // Причина снята и источник можно сбросить
	xRejected         : BOOL; // Одноцикловый признак отклонённого запроса
	udiRejectSequence : UDINT; // Счётчик отклонённых запросов для надёжного чтения HMI
END_STRUCT
END_TYPE

// Device/Application/ST/ST_POINT/E_POINT_NAME
{attribute 'qualified_only'}
{attribute 'strict'}
TYPE E_POINT_NAME :
(	
	NONE,
	MACHINE_1_ABOVE,
	MACHINE_1_INSIDE, // Legacy: исключена из редактора, сохранена ради числового протокола
	MACHINE_1_CHUCK_APROACH,
	MACHINE_1_CHUCK_POSITION,
	MACHINE_2_ABOVE,
	MACHINE_2_INSIDE, // Legacy: исключена из редактора, сохранена ради числового протокола
	MACHINE_2_CHUCK_APROACH,
	MACHINE_2_CHUCK_POSITION,
	MACHINE_3_ABOVE,
	MACHINE_3_INSIDE, // Legacy: исключена из редактора, сохранена ради числового протокола
	MACHINE_3_CHUCK_APROACH,
	MACHINE_3_CHUCK_POSITION,
	MAGAZINE_DETAIL,
	MAGAZINE_TAKE_DETAIL,
	MAGAZINE_PUT_DETAIL,
	MAGAZINE_CHANGE_DETAIL,
	HOME_SAFETY,
	MAGAZINE_RETURN_BLANK, // Legacy: сохранено только ради прежнего числового значения
	MAGAZINE_SAFE, // Безопасная точка над активным слотом
	MAGAZINE_IN_SLOT, // Рабочая точка внутри активного слота
	MAGAZINE_CHANGE, // Безопасная точка переворота над активным слотом
	MAGAZINE_1_DETAIL, // Базовая точка рабочей зоны первого магазина
	MAGAZINE_2_DETAIL, // Базовая точка рабочей зоны второго магазина
	GEOMETRY_1_PLACE,
	GEOMETRY_1_SAFE,
	GEOMETRY_1_CHANGE,
	GEOMETRY_2_PLACE,
	GEOMETRY_2_SAFE,
	GEOMETRY_2_CHANGE

);
END_TYPE

// Device/Application/ST/ST_CELL/ST_CELL_SAFETY_FAULT_REQUEST
TYPE ST_CELL_SAFETY_FAULT_REQUEST :
STRUCT
	xEnabled : BOOL; // Общее разрешение диагностических инъекций
	axEmergencyStopStation : ARRAY [1..4] OF BOOL;
	axEmergencyStopCabinet : ARRAY [1..2] OF BOOL;
	xEmergencyStopMpg      : BOOL;
	xPhaseRelayFault       : BOOL;
	xPressureRelayFault    : BOOL;
	xSafetyRelayFault      : BOOL;
	axDoorUnlocked         : ARRAY [1..4] OF BOOL;
END_STRUCT
END_TYPE

// Device/Application/ST/ST_MAGAZINE/ST_MAGAZINE_HMI_COMMAND
TYPE ST_MAGAZINE_HMI_COMMAND :
STRUCT
	{attribute 'symbol' := 'read'}
	xEnable : BOOL; // Импульс включения технологической логики магазина
	{attribute 'symbol' := 'read'}
	xDisable : BOOL; // Импульс отключения технологической логики магазина
	{attribute 'symbol' := 'read'}
	xStop : BOOL; // Остановить выполняемую операцию магазина
	{attribute 'symbol' := 'read'}
	xReset : BOOL; // Сброс ошибок магазина
	{attribute 'symbol' := 'read'}
	xFill : BOOL; // Заполнить кассету заготовками по текущей карте типов
	{attribute 'symbol' := 'read'}
	xClear : BOOL; // Полностью очистить кассету
	xCycleSlot : BOOL; // Переключить содержимое выбранного слота
	{attribute 'symbol' := 'read'}
	xApplySlot : BOOL; // Явно записать состояние и тип выбранного слота
	{attribute 'symbol' := 'read'}
	xApplyPitchX : BOOL; // Применить новый шаг слотов по X
	{attribute 'symbol' := 'read'}
	xApplyPitchY : BOOL; // Применить новый шаг слотов по Y
	uiEditSlot : UINT; // Слот кассеты, 1..120
	uiEditDetailType : UINT; // 0=NONE, 1=BLANK, 2=DETAIL
	uiEditProductType : UINT; // Тип изделия 1..3; для NONE игнорируется
	lrEditPitchX : LREAL; // Запрошенный шаг слотов по X
	lrEditPitchY : LREAL; // Запрошенный шаг слотов по Y
END_STRUCT
END_TYPE

// Device/Application/ST/ST_MAGAZINE/ST_TWO_PALLET_STATUS
TYPE ST_TWO_PALLET_STATUS :
STRUCT
	uiStep : UINT;
	uiFaultStep : UINT; // Шаг, на котором появился последний новый аварийный бит
	uiCandidate : UINT; // Расстановка, совместимая с датчиками; не измерение палет
	uiRobotPallet : UINT := 1; // Учётный номер, меняется только после подтверждения/завершения обмена
	uiSelected : UINT;
	udiRevision : UDINT;
	xEnabled : BOOL;
	xConfirmed : BOOL;
	xReady : BOOL;
	xBusy : BOOL;
	xError : BOOL;
	xHomeRequired : BOOL;
	xConfigValid : BOOL;
	xConfirmAllowed : BOOL;
	xStartAllowed : BOOL;
	xEnableAllowed : BOOL;
	xSwapAllowed : BOOL;
	xPowerAllowed : BOOL;
	xDriveResetAllowed : BOOL;
	xHomeAllowed : BOOL;
	xLowerAllowed : BOOL;
	xRaiseAllowed : BOOL;
	xSelectAllowed : BOOL;
	xLockAllowed : BOOL;
	xStopAllowed : BOOL;
	xMoveAllowed : BOOL;
	xJogAllowed : BOOL;
	xTeachOperatorAllowed : BOOL;
	xTeachWorkAllowed : BOOL;
	xResetAllowed : BOOL;
	xEditAllowed : BOOL;
	xEdit1Allowed : BOOL;
	xEdit2Allowed : BOOL;
	xLoadAllowed : BOOL; // Подтвердить загрузку текущей операторской палеты
	xConfigAllowed : BOOL;
	xCompleted : BOOL;
	xCommandAccepted : BOOL;
	uiReason : UINT;
	dwError : DWORD;
	stWarning : ST_WARNING_EVENT;
	Input : ST_TWO_PALLET_INPUT;
	rP1 : REAL; // Оценка нормализованного положения для 3D, не датчик палеты
	rP2 : REAL;
	rLift : REAL;
	xAutoSwapEnabled : BOOL; // Настройка автоматической смены палет
END_STRUCT
END_TYPE

// Device/Application/ST/ST_MAGAZINE/ST_TWO_PALLET_STORE
TYPE ST_TWO_PALLET_STORE :
STRUCT
	astPallet : ARRAY [1..2] OF ST_MAGAZINE_INVENTORY;
	axLoaded : ARRAY [1..2] OF BOOL; // Снимается после обмена и каждого редактирования
END_STRUCT
END_TYPE

// Device/Application/ST/ST_GRIPPER/ST_GRIPPER_ERROR
TYPE ST_GRIPPER_ERROR :
STRUCT
	GRIPPER_1_ERROR : BOOL; // Ошибка первого захвата
	GRIPPER_2_ERROR : BOOL; // Ошибка второго захвата
	ROTATION_ERROR  : BOOL; // Ошибка механизма поворота
	ACTION_ERROR    : BOOL; // Получено недопустимое действие
	GLOBAL_ERROR    : BOOL; // Глобальная ошибка симуляции захвата
END_STRUCT
END_TYPE

// Device/Application/ST/ST_AXIS/ST_AXIS_ERROR
TYPE ST_AXIS_ERROR :
STRUCT
	MC_POWER_ERROR       : BOOL; // Ошибка MC_Power
	MC_RESET_ERROR       : BOOL; // Ошибка MC_Reset
	MC_STOP_ERROR        : BOOL; // Ошибка MC_Stop
	MC_JOG_ERROR         : BOOL; // Ошибка MC_Jog
	MC_HOME_ERROR        : BOOL; // Ошибка MC_Home
	MC_MOVE_ABS_ERROR    : BOOL; // Ошибка MC_MoveAbsolute
	MC_MOVE_REL_ERROR    : BOOL; // Ошибка MC_MoveRelative
	READ_POSITION_ERROR  : BOOL; // Ошибка чтения позиции
	READ_STATUS_ERROR    : BOOL; // Ошибка чтения статуса оси
	AXIS_ERRORSTOP       : BOOL; // Ось находится в ErrorStop
	FB_ERROR_OCCURRED    : BOOL; // SoftMotion сообщил внутреннюю ошибку
	COMMAND_ABORTED      : BOOL; // Команда движения была прервана
	UNKNOWN_AXIS_ERROR   : BOOL; // Неизвестная ошибка оси
	DRIVE_AXIS_ERROR     : BOOL; // Ошибка привода оси
	POWER_FEEDBACK_LOST  : BOOL; // Потеря силовой готовности при активной команде питания
	POWER_PERMIT_LOST    : BOOL; // Потеря разрешения питания
	GLOBAL_DURING_POWER  : BOOL; // Глобальная ошибка при включении
	GLOBAL_DURING_READY  : BOOL; // Глобальная ошибка в готовности
	GLOBAL_DURING_MOTION : BOOL; // Глобальная ошибка во время движения
	JOG_CONFLICT         : BOOL; // Одновременно поданы Jog+ и Jog-
	MOVE_ABS_NOT_HOMED   : BOOL; // Абсолютное движение без Home
	MOVE_REL_NOT_HOMED   : BOOL; // Относительное движение без Home
	STEP_TIMEOUT         : BOOL; // Превышено время выполнения шага
	UNKNOWN_STEP         : BOOL; // Неизвестное состояние автомата
END_STRUCT
END_TYPE

// Device/Application/ST/ST_MAGAZINE/E_MAGAZINE_OPERATION
{attribute 'qualified_only'}
{attribute 'strict'}
TYPE E_MAGAZINE_OPERATION :
(
	NONE         := 0,
	PUT          := 1,
	TAKE         := 2,
	CHANGE       := 3,
	RETURN_BLANK := 4
);
END_TYPE

// Device/Application/ST/ST_MACHINE/ST_MACHINE_IO_STATUS
TYPE ST_MACHINE_IO_STATUS :
STRUCT
	xReady          : BOOL; // Станок готов принимать команды
	xAlarm          : BOOL; // Активна авария станка
	xDoorOpen       : BOOL; // Роботный люк открыт; имя сохранено для совместимости
	xDoorClosed     : BOOL; // Роботный люк закрыт; имя сохранено для совместимости
	xHatchLocked    : BOOL; // Замок роботного люка закрыт (0 — открыт, 1 — закрыт)
	xSafetyDoorOpen   : BOOL; // Операторская дверь открыта
	xSafetyDoorClosed : BOOL; // Операторская дверь закрыта
	xChuckClamped   : BOOL; // Патрон зажат
	xChuckUnclamped : BOOL; // Патрон разжат
	xCycleActive    : BOOL; // Выполняется цикл обработки
	xCycleDone      : BOOL; // Цикл обработки завершён
	tRemaining      : TIME; // Оставшееся время обработки
END_STRUCT
END_TYPE

// Device/Application/ST/ST_MAGAZINE/ST_MAGAZINE_INVENTORY
TYPE ST_MAGAZINE_INVENTORY :
STRUCT
	aSlots : ARRAY [1..GVL_CELL_SETTINGS.MagazineSlots] OF ST_DETAIL; // Единственная статичная кассета
END_STRUCT
END_TYPE

// Device/Application/ST/ST_ROBOT/E_ROBOT_CONTROL_MODE
{attribute 'qualified_only'}
{attribute 'strict'}
TYPE E_ROBOT_CONTROL_MODE :
(
	SOFTMOTION := 0,
	MODBUS_TCP := 1
);
END_TYPE

// Device/Application/ST/ST_MACHINE/E_MACHINE_POINTS
{attribute 'qualified_only'}
{attribute 'strict'}
TYPE E_MACHINE_POINTS :
(
	NONE,     
	ABOVE,         
    INSIDE,        
    CHUCK_APPROACH, 
    CHUCK         
);
END_TYPE

// Device/Application/ST/ST_AXIS/ST_AXIS_COMMANDS
TYPE ST_AXIS_COMMANDS :
STRUCT
    xEnable            : BOOL; // Импульс запроса включения оси
    xDisable           : BOOL; // Импульс запроса отключения оси
	xGlobalError       : BOOL; // Глобальная ошибка ячейки
	xPowerPermit       : BOOL; // Разрешение подачи питания на привод
    xResetAllError     : BOOL; // Общий сброс ошибок оси
    xResetAxisError    : BOOL; // Сброс ошибок привода и SoftMotion
    xResetLogicalError : BOOL; // Сброс логических ошибок блока
    xStop              : BOOL; // Команда контролируемой остановки
    xHome              : BOOL; // Команда поиска домашней позиции
    xMoveAbsolute      : BOOL; // Команда абсолютного перемещения
    xMoveRelative      : BOOL; // Команда относительного перемещения
    xJogPositive       : BOOL; // Толчковое движение в положительном направлении
    xJogNegative       : BOOL; // Толчковое движение в отрицательном направлении
END_STRUCT
END_TYPE

// Device/Application/ST/ST_MAGAZINE/ST_TWO_PALLET_REQUEST
TYPE ST_TWO_PALLET_REQUEST :
STRUCT
	uiMagazine : UINT; // 0: конфигурация линии; 1..2: отдельный магазин
	uiCommand : UINT;
	uiValue : UINT;
	uiSlot : UINT;
	uiContent : UINT;
	uiProductType : UINT;
	udiRevision : UDINT;
	Config : ST_TWO_PALLET_CONFIG;
END_STRUCT
END_TYPE

// Device/Application/ST/ST_GEOMETRY_CONTROL/ST_GEOMETRY_EVENT
TYPE ST_GEOMETRY_EVENT :
STRUCT
	udiSequence : UDINT;
	udiTimeMs : UDINT; // Монотонные часы PLC, не настенные часы
	uiEnvironment : UINT; // NORMAL=0, SIMULATION=1, SC500_BENCH=2
	Call : ST_GEOMETRY_CALL;
END_STRUCT
END_TYPE

// Device/Application/ST/ST_MAGAZINE/ST_TWO_PALLET_OUTPUT
TYPE ST_TWO_PALLET_OUTPUT :
STRUCT
	xLiftUp : BOOL;
	xLiftDown : BOOL;
	xLockOut : BOOL;
	xLockIn : BOOL;
	xStopOut : BOOL;
	xStopIn : BOOL;
	xPowerOn : BOOL;
	xPowerOff : BOOL;
	xDriveReset : BOOL;
	xHome : BOOL;
	xMove : BOOL;
	xStop : BOOL;
	xJogPositive : BOOL;
	xJogNegative : BOOL;
	xTeachOperator : BOOL;
	xTeachWork : BOOL;
	lrTarget : LREAL;
END_STRUCT
END_TYPE

// Device/Application/ST/ST_MOTION_MANAGER/ST_MOTION_MANAGER_STATUS
TYPE ST_MOTION_MANAGER_STATUS :
STRUCT
	xReady        : BOOL; // Менеджер готов принять команду
	xBusy         : BOOL; // Выполняется движение
	xDone         : BOOL; // Движение завершено
	xError        : BOOL; // Менеджер находится в ошибке
	eCurrentPoint : E_POINT_NAME; // Последняя достигнутая точка
END_STRUCT
END_TYPE

